(* IEC 61131-3 sources: daoli-st-library/DL_Device (part 10) *)

(* ---- FC_DL_RefSatPressToTemp.st ---- *)
(*
  ============================================================
  组件名 : FC_DL_RefSatPressToTemp
  分类   : DL_Device
  功能   : 制冷剂饱和压力转饱和温度，内置 R134a 与 R410A 分段线性表并做区间插值
  开源溯源 : internal-design（本轮无外部代码逐行引用）
             参考语义 : 无外部参考
  复杂度 : C2
  版本   : 1.0.0
  ============================================================
  表口径 : 压力为绝对压力 [bar abs]，温度为 [摄氏度]，两行表按 R134a 与 R410A 顺序平铺，
           行内压力严格升序；压力越出表范围时取端点温度并置 bValid 为假。
*)

FUNCTION FC_DL_RefSatPressToTemp : REAL
VAR_INPUT
    rPressBarA    : REAL; // 饱和绝对压力 [bar abs] saturation absolute pressure [bar abs]
    nRefrigerant  : INT; // 制冷剂 1=R134a 2=R410A [代号] refrigerant 1 for R134a and 2 for R410A [code]
END_VAR
VAR_OUTPUT
    rTempC : REAL; // 饱和温度 [摄氏度] saturation temperature [degree celsius]
    bValid : BOOL; // 结果有效标志 result validity flag
END_VAR
VAR CONSTANT
    afPress : ARRAY[0..1, 0..7] OF REAL := [1.0, 2.0, 4.0, 6.0, 8.0, 10.0, 14.0, 18.0, 1.0, 2.0, 4.0, 6.0, 8.0, 10.0, 14.0, 18.0]; // 饱和压力表 [bar abs] saturation pressure table [bar abs]
    afTemp  : ARRAY[0..1, 0..7] OF REAL := [-26.1, -10.1, 8.9, 21.6, 31.3, 39.4, 52.4, 62.5, -51.4, -34.1, -14.1, 0.4, 11.4, 20.5, 34.4, 45.0]; // 饱和温度表 [摄氏度] saturation temperature table [degree celsius]
    DL_IDX_LAST : INT := 7; // 表末下标 last table index
    DL_EPS_R    : REAL := 1.0E-6; // 实数零判定阈值 real zero threshold
END_VAR
VAR
    nRow  : INT := 0; // 表行号 0=R134a 1=R410A [行] table row number [row]
    nSeg  : INT := -1; // 命中区间下标，负为未命中 [段] hit segment index, negative when missing [segment]
    i     : INT := 0; // 区间游标 [段] segment cursor [segment]
    _rSpan: REAL := 0.0; // 区间压力跨度 [bar] segment pressure span [bar]
    _rFrac: REAL := 0.0; // 区间插值比例 [无量纲] interpolation fraction [dimensionless]
    _rT   : REAL := 0.0; // 温度中间量 [摄氏度] intermediate temperature [degree celsius]
END_VAR

// 段 1｜出口预置 preset the exit
FC_DL_RefSatPressToTemp := 0.0; // 缺省返回零 default zero return
rTempC := 0.0; // 温度预置零 temperature preset to zero
bValid := FALSE; // 计算完成前不认结果 unusable before the calculation
// 段 2｜非有限闸与制冷剂代号闸 finiteness gate and refrigerant code gate
IF (rPressBarA <> rPressBarA) OR (nRefrigerant < 1) OR (nRefrigerant > 2) THEN
    RETURN; // 非有限或代号非法即无效 non finite or an illegal code is void
END_IF
nRow := nRefrigerant - 1; // 行号由代号减一得出 the row index is the code minus one
// 段 3｜区间搜索 segment search over the ascending pressure table
FOR i := 0 TO (DL_IDX_LAST - 1) DO
    IF (rPressBarA >= afPress[nRow, i]) AND (rPressBarA <= afPress[nRow, i + 1]) THEN
        nSeg := i; // 命中升序区间 a segment is hit
    END_IF
END_FOR
// 段 4｜越界端点处理 endpoint handling for the out of table pressures
IF nSeg < 0 THEN
    IF rPressBarA < afPress[nRow, 0] THEN
        rTempC := afTemp[nRow, 0]; // 低于表底取表首温度 a pressure below the table takes the first temperature
    ELSE
        rTempC := afTemp[nRow, DL_IDX_LAST]; // 高于表顶取表末温度 a pressure above the table takes the last temperature
    END_IF
    RETURN; // 越界置无效并输出端点值 the out of table case is void with the endpoint emitted
END_IF
// 段 5｜线性插值 linear interpolation inside the hit segment
_rSpan := afPress[nRow, nSeg + 1] - afPress[nRow, nSeg]; // 区间压力跨度 segment pressure span
IF ABS(_rSpan) < DL_EPS_R THEN
    RETURN; // 跨度近零无法插值 a near zero span cannot interpolate
END_IF
_rFrac := (rPressBarA - afPress[nRow, nSeg]) / _rSpan; // 区间内插值比例 the fraction inside the segment
_rT := afTemp[nRow, nSeg] + _rFrac * (afTemp[nRow, nSeg + 1] - afTemp[nRow, nSeg]); // 端点温度线性插值 linear blend of the two temperatures
rTempC := _rT; // 温度落定 land the temperature
bValid := TRUE; // 结果可用 result usable
FC_DL_RefSatPressToTemp := _rT; // 函数返回饱和温度 return the saturation temperature
END_FUNCTION

(* ---- FC_DL_RefSatTempToPress.st ---- *)
(*
  ============================================================
  组件名 : FC_DL_RefSatTempToPress
  分类   : DL_Device
  功能   : 制冷剂饱和温度转饱和压力，内置 R134a 与 R410A 分段线性表并做区间插值
  开源溯源 : internal-design（本轮无外部代码逐行引用）
             参考语义 : 无外部参考
  复杂度 : C2
  版本   : 1.0.0
  ============================================================
  表口径 : 与压力查温度件同源的两张表，按温度升序重排后以温度为自变量插值压力；
           温度为绝对压力 [bar abs] 输出，温度越出表范围时取端点压力并置 bValid 为假。
*)

FUNCTION FC_DL_RefSatTempToPress : REAL
VAR_INPUT
    rTempC       : REAL; // 饱和温度 [摄氏度] saturation temperature [degree celsius]
    nRefrigerant : INT; // 制冷剂 1=R134a 2=R410A [代号] refrigerant 1 for R134a and 2 for R410A [code]
END_VAR
VAR_OUTPUT
    rPressBarA : REAL; // 饱和绝对压力 [bar abs] saturation absolute pressure [bar abs]
    bValid     : BOOL; // 结果有效标志 result validity flag
END_VAR
VAR CONSTANT
    afTemp  : ARRAY[0..1, 0..7] OF REAL := [-26.1, -10.1, 8.9, 21.6, 31.3, 39.4, 52.4, 62.5, -51.4, -34.1, -14.1, 0.4, 11.4, 20.5, 34.4, 45.0]; // 饱和温度表，行内升序 [摄氏度] saturation temperature table ascending inside each row [degree celsius]
    afPress : ARRAY[0..1, 0..7] OF REAL := [1.0, 2.0, 4.0, 6.0, 8.0, 10.0, 14.0, 18.0, 1.0, 2.0, 4.0, 6.0, 8.0, 10.0, 14.0, 18.0]; // 饱和压力表 [bar abs] saturation pressure table [bar abs]
    DL_IDX_LAST : INT := 7; // 表末下标 last table index
    DL_EPS_R    : REAL := 1.0E-6; // 实数零判定阈值 real zero threshold
END_VAR
VAR
    nRow  : INT := 0; // 表行号 0=R134a 1=R410A [行] table row number [row]
    nSeg  : INT := -1; // 命中区间下标，负为未命中 [段] hit segment index, negative when missing [segment]
    i     : INT := 0; // 区间游标 [段] segment cursor [segment]
    _rSpan: REAL := 0.0; // 区间温度跨度 [K] segment temperature span [kelvin]
    _rFrac: REAL := 0.0; // 区间插值比例 [无量纲] interpolation fraction [dimensionless]
    _rP   : REAL := 0.0; // 压力中间量 [bar abs] intermediate pressure [bar abs]
END_VAR

// 段 1｜出口预置 preset the exit
FC_DL_RefSatTempToPress := 0.0; // 缺省返回零 default zero return
rPressBarA := 0.0; // 压力预置零 pressure preset to zero
bValid := FALSE; // 计算完成前不认结果 unusable before the calculation
// 段 2｜非有限闸与制冷剂代号闸 finiteness gate and refrigerant code gate
IF (rTempC <> rTempC) OR (nRefrigerant < 1) OR (nRefrigerant > 2) THEN
    RETURN; // 非有限或代号非法即无效 non finite or an illegal code is void
END_IF
nRow := nRefrigerant - 1; // 行号由代号减一得出 the row index is the code minus one
// 段 3｜区间搜索 segment search over the ascending temperature table
FOR i := 0 TO (DL_IDX_LAST - 1) DO
    IF (rTempC >= afTemp[nRow, i]) AND (rTempC <= afTemp[nRow, i + 1]) THEN
        nSeg := i; // 命中升序区间 a segment is hit
    END_IF
END_FOR
// 段 4｜越界端点处理 endpoint handling for the out of table temperatures
IF nSeg < 0 THEN
    IF rTempC < afTemp[nRow, 0] THEN
        rPressBarA := afPress[nRow, 0]; // 低于表底取表首压力 a temperature below the table takes the first pressure
    ELSE
        rPressBarA := afPress[nRow, DL_IDX_LAST]; // 高于表顶取表末压力 a temperature above the table takes the last pressure
    END_IF
    RETURN; // 越界置无效并输出端点值 the out of table case is void with the endpoint emitted
END_IF
// 段 5｜线性插值 linear interpolation inside the hit segment
_rSpan := afTemp[nRow, nSeg + 1] - afTemp[nRow, nSeg]; // 区间温度跨度 segment temperature span
IF ABS(_rSpan) < DL_EPS_R THEN
    RETURN; // 跨度近零无法插值 a near zero span cannot interpolate
END_IF
_rFrac := (rTempC - afTemp[nRow, nSeg]) / _rSpan; // 区间内插值比例 the fraction inside the segment
_rP := afPress[nRow, nSeg] + _rFrac * (afPress[nRow, nSeg + 1] - afPress[nRow, nSeg]); // 端点压力线性插值 linear blend of the two pressures
rPressBarA := _rP; // 压力落定 land the pressure
bValid := TRUE; // 结果可用 result usable
FC_DL_RefSatTempToPress := _rP; // 函数返回饱和压力 return the saturation pressure
END_FUNCTION

(* ---- FC_DL_RefSubcoolCalc.st ---- *)
(*
  ============================================================
  组件名 : FC_DL_RefSubcoolCalc
  分类   : DL_Device
  功能   : 液管过冷度计算，由冷凝饱和温度与液管温度求过冷度并分档判定
  开源溯源 : internal-design（本轮无外部代码逐行引用）
             参考语义 : 无外部参考
  复杂度 : C1
  版本   : 1.0.0
  ============================================================
*)

FUNCTION FC_DL_RefSubcoolCalc : REAL
VAR_INPUT
    rLiquidTempC    : REAL; // 液管实测温度 [摄氏度] measured liquid line temperature [degree celsius]
    rSatLiquidTempC : REAL; // 液管饱和温度 [摄氏度] saturation temperature at the liquid pressure [degree celsius]
    rScLow          : REAL; // 过冷度下限 [K] lower subcooling bound [kelvin]
    rScHigh         : REAL; // 过冷度上限 [K] upper subcooling bound [kelvin]
END_VAR
VAR_OUTPUT
    rSubcoolK : REAL; // 液管过冷度 [K] liquid subcooling [kelvin]
    nStatus   : INT; // 分档 0正常 1偏低 2偏高 [档] status 0 normal, 1 low, 2 high [band]
    bValid    : BOOL; // 结果有效标志 result validity flag
END_VAR
VAR
    _bFin  : BOOL := FALSE; // 四输入有限性判定 finiteness verdict of the four inputs
    _rSc   : REAL := 0.0; // 过冷度中间量 [K] intermediate subcooling [kelvin]
    _rLo   : REAL := 0.0; // 钳位后的下限 [K] clamped lower bound [kelvin]
    _rHi   : REAL := 0.0; // 钳位后的上限 [K] clamped upper bound [kelvin]
END_VAR

// 段 1｜出口预置 preset the exit
FC_DL_RefSubcoolCalc := 0.0; // 缺省返回零 default zero return
rSubcoolK := 0.0; // 过冷度预置零 subcooling preset to zero
nStatus := 0; // 分档预置正常 status preset normal
bValid := FALSE; // 计算完成前不认结果 unusable before the calculation
// 段 2｜非有限闸 finiteness gate
_bFin := (rLiquidTempC = rLiquidTempC) AND (rSatLiquidTempC = rSatLiquidTempC) AND (rScLow = rScLow) AND (rScHigh = rScHigh); // 四输入自反判定 self comparison of the four inputs
IF NOT _bFin THEN
    RETURN; // 非有限即无效 non finite means invalid
END_IF
// 段 3｜主体过冷度 main subcooling，口径为饱和温度减液管温度 saturation minus the liquid temperature
_rSc := rSatLiquidTempC - rLiquidTempC; // 饱和温度减液管温度 saturation minus the liquid temperature
rSubcoolK := _rSc; // 过冷度落定 land the subcooling
// 段 4｜上下限整形 bound reshape
_rLo := rScLow; // 取下限 take the lower bound
_rHi := rScHigh; // 取上限 take the upper bound
IF _rLo > _rHi THEN
    _rLo := rScHigh; // 上下限倒置时下限取原上限 an inverted pair swaps the lower bound
    _rHi := rScLow; // 上下限倒置时上限取原下限 an inverted pair swaps the upper bound
END_IF
// 段 5｜双向分档判定 directional status verdict
IF _rSc < _rLo THEN
    nStatus := 1; // 过冷度偏低 subcooling too low
ELSIF _rSc > _rHi THEN
    nStatus := 2; // 过冷度偏高 subcooling too high
ELSE
    nStatus := 0; // 区间内正常 inside the normal band
END_IF
bValid := TRUE; // 结果可用 result usable
FC_DL_RefSubcoolCalc := _rSc; // 函数返回过冷度 return the subcooling
END_FUNCTION

(* ---- FC_DL_RefSuperheatCalc.st ---- *)
(*
  ============================================================
  组件名 : FC_DL_RefSuperheatCalc
  分类   : DL_Device
  功能   : 吸气过热度计算，由吸气温度与对应饱和温度求过热度并分档判定
  开源溯源 : internal-design（本轮无外部代码逐行引用）
             参考语义 : 无外部参考
  复杂度 : C1
  版本   : 1.0.0
  ============================================================
*)

FUNCTION FC_DL_RefSuperheatCalc : REAL
VAR_INPUT
    rSuctionTempC    : REAL; // 吸气实测温度 [摄氏度] measured suction temperature [degree celsius]
    rSatSuctionTempC : REAL; // 吸气饱和温度 [摄氏度] saturation temperature at the suction pressure [degree celsius]
    rShLow           : REAL; // 过热度下限 [K] lower superheat bound [kelvin]
    rShHigh          : REAL; // 过热度上限 [K] upper superheat bound [kelvin]
END_VAR
VAR_OUTPUT
    rSuperheatK : REAL; // 吸气过热度 [K] suction superheat [kelvin]
    nStatus     : INT; // 分档 0正常 1偏低 2偏高 [档] status 0 normal, 1 low, 2 high [band]
    bValid      : BOOL; // 结果有效标志 result validity flag
END_VAR
VAR
    _bFin  : BOOL := FALSE; // 四输入有限性判定 finiteness verdict of the four inputs
    _rSh   : REAL := 0.0; // 过热度中间量 [K] intermediate superheat [kelvin]
    _rLo   : REAL := 0.0; // 钳位后的下限 [K] clamped lower bound [kelvin]
    _rHi   : REAL := 0.0; // 钳位后的上限 [K] clamped upper bound [kelvin]
END_VAR

// 段 1｜出口预置 preset the exit
FC_DL_RefSuperheatCalc := 0.0; // 缺省返回零 default zero return
rSuperheatK := 0.0; // 过热度预置零 superheat preset to zero
nStatus := 0; // 分档预置正常 status preset normal
bValid := FALSE; // 计算完成前不认结果 unusable before the calculation
// 段 2｜非有限闸 finiteness gate
_bFin := (rSuctionTempC = rSuctionTempC) AND (rSatSuctionTempC = rSatSuctionTempC) AND (rShLow = rShLow) AND (rShHigh = rShHigh); // 四输入自反判定 self comparison of the four inputs
IF NOT _bFin THEN
    RETURN; // 非有限即无效 non finite means invalid
END_IF
// 段 3｜主体过热度 main superheat
_rSh := rSuctionTempC - rSatSuctionTempC; // 吸气温度减饱和温度 suction minus saturation
rSuperheatK := _rSh; // 过热度落定 land the superheat
// 段 4｜上下限整形 bound reshape
_rLo := rShLow; // 取下限 take the lower bound
_rHi := rShHigh; // 取上限 take the upper bound
IF _rLo > _rHi THEN
    _rLo := rShHigh; // 上下限倒置时下限取原上限 an inverted pair swaps the lower bound
    _rHi := rShLow; // 上下限倒置时上限取原下限 an inverted pair swaps the upper bound
END_IF
// 段 5｜双向分档判定 directional status verdict
IF _rSh < _rLo THEN
    nStatus := 1; // 过热度偏低 superheat too low
ELSIF _rSh > _rHi THEN
    nStatus := 2; // 过热度偏高 superheat too high
ELSE
    nStatus := 0; // 区间内正常 inside the normal band
END_IF
bValid := TRUE; // 结果可用 result usable
FC_DL_RefSuperheatCalc := _rSh; // 函数返回过热度 return the superheat
END_FUNCTION

(* ---- FC_DL_SheetPeelForceCalc.st ---- *)
(*
  ============================================================
  组件名 : FC_DL_SheetPeelForceCalc
  分类   : DL_Device
  功能   : 片材剥离力计算，由接触面积粘附强度与静电电压求剥离力并按剥离角折减
  复杂度 : C2
  版本   : 1.0.0
  作者   : 道莅工业代码库工厂 / R81
  日期   : 2026-11-24
  开源溯源 : clean-room（no upstream）—— 依据公开工程公式自研，未复制任何上游实现
  红线自检 : R1 无GVL/R2 无物理地址/R3 纯IEC/R4 防除零/R5 双语注释
  接口说明 :
      粘附分量 = 接触面积(m2) * 粘附强度(Pa)，面积由 mm2 乘 1e-6，强度由 kPa 乘 1000。
      静电分量 = 静电电压(kV) * 0.05，系数为工程经验折算，单位 N/kV。
      剥离角修正系数 = (1 + COS(角度)) / 2，归一到 0 度时为 1、90 度为 0.5、180 度为 0，便于跨机型比较。
      剥离力超过 50 N 判需要外部辅助剥离。
  ============================================================
*)
FUNCTION FC_DL_SheetPeelForceCalc : BOOL
VAR_INPUT
    bEnable       : BOOL; // 使能：TRUE 时计算 / Enable: TRUE to compute
    bErr          : BOOL; // 外部故障：TRUE 时立即退出并置结果无效 / External fault: TRUE aborts with invalid result
    rArea_mm2     : REAL; // 片材与承载面接触面积 [mm2] / contact area between sheet and support [square millimetre]
    rAdhesion_kpa : REAL; // 单位面积粘附强度 [kPa] / adhesion strength per unit area [kilopascal]
    rStaticKv     : REAL; // 片材静电电位 [kV] / electrostatic potential of the sheet [kilovolt]
    rPeelAngleDeg : REAL; // 剥离角度，0 度表示垂直拉起 [度] / peel angle, zero means lifting perpendicular [degree]
END_VAR
VAR_OUTPUT
    rAdhesionN : REAL; // 粘附力分量 [N] / adhesion force component [newton]
    rStaticN   : REAL; // 静电力分量 [N] / electrostatic force component [newton]
    rAngleFactor : REAL; // 剥离角折减系数，0~1 [无量纲] / peel angle reduction factor from 0 to 1 [dimensionless]
    rPeelN     : REAL; // 综合剥离力 [N] / resultant peel force [newton]
    bNeedAssist : BOOL; // 需要辅助：TRUE 表示剥离力超过 50 N / assistance required, TRUE when the peel force exceeds 50 newton
    bValid     : BOOL; // 输出有效：TRUE 表示结果可用 / Output valid
END_VAR
VAR CONSTANT
    DL_R_MAX     : REAL := 3.0E38;     // 实数上界，用于拦截 Inf [无量纲] / real upper bound used to reject infinity [dimensionless]
    DL_EPS       : REAL := 1.0E-12;    // 除零判定阈值 [无量纲] / division guard threshold [dimensionless]
    DL_MM2_TO_M2 : REAL := 1.0E-6;     // 平方毫米折平方米系数 [m2/mm2] / square millimetre to square metre factor [square metre per square millimetre]
    DL_KPA_TO_PA : REAL := 1000.0;     // 千帕折帕系数 [Pa/kPa] / kilopascal to pascal factor [pascal per kilopascal]
    DL_KV_TO_N   : REAL := 0.05;       // 每千伏静电折算力 [N/kV] / electrostatic force per kilovolt [newton per kilovolt]
    DL_DEG_TO_RAD : REAL := 0.0174533; // 度转弧度系数 [rad/度] / degree to radian factor [radian per degree]
    DL_HALF      : REAL := 0.5;        // 二分之一，用于角度系数归一 [无量纲] / one half used to normalise the angle factor [dimensionless]
    DL_ONE       : REAL := 1.0;        // 单位常量 [无量纲] / unity constant [dimensionless]
    DL_ASSIST_N  : REAL := 50.0;       // 辅助剥离门限 [N] / assistance threshold [newton]
    DL_ANGLE_MAX : REAL := 180.0;      // 剥离角允许上限 [度] / permitted upper bound of the peel angle [degree]
    DL_STAT_MAX  : REAL := 1000.0;     // 静电电位合理上限 [kV] / sanity upper bound of the electrostatic potential [kilovolt]
END_VAR
VAR
    _bFin  : BOOL := FALSE; // 输入有限性判定结果 / input finiteness verdict
    _rRad  : REAL := 0.0;   // 剥离角折算弧度 [rad] / peel angle in radian [radian]
END_VAR

    // 段 1｜出口预置
    rAdhesionN := 0.0;
    rStaticN := 0.0;
    rAngleFactor := 0.0;
    rPeelN := 0.0;
    bNeedAssist := FALSE;
    bValid := FALSE;
    // 段 2｜使能闸与外部故障闸
    IF NOT bEnable THEN
        RETURN;
    END_IF;
    IF bErr THEN
        RETURN;
    END_IF;
    // 段 3｜非有限闸
    _bFin := (rArea_mm2 = rArea_mm2) AND (ABS(rArea_mm2) <= DL_R_MAX) AND (rAdhesion_kpa = rAdhesion_kpa) AND (ABS(rAdhesion_kpa) <= DL_R_MAX) AND (rStaticKv = rStaticKv) AND (ABS(rStaticKv) <= DL_R_MAX) AND (rPeelAngleDeg = rPeelAngleDeg) AND (ABS(rPeelAngleDeg) <= DL_R_MAX);
    IF NOT _bFin THEN
        RETURN;
    END_IF;
    // 段 4｜域闸：面积非负、粘附强度非负、静电位非负且合理、角度 0~180
    IF (rArea_mm2 < 0.0) OR (rAdhesion_kpa < 0.0) OR (rStaticKv < 0.0) OR (rStaticKv > DL_STAT_MAX) THEN
        RETURN;
    END_IF;
    IF (rPeelAngleDeg < 0.0) OR (rPeelAngleDeg > DL_ANGLE_MAX) THEN
        RETURN;
    END_IF;
    // 段 5｜两个力分量
    rAdhesionN := rArea_mm2 * DL_MM2_TO_M2 * rAdhesion_kpa * DL_KPA_TO_PA;
    rStaticN := rStaticKv * DL_KV_TO_N;
    // 段 6｜角度折减系数
    _rRad := rPeelAngleDeg * DL_DEG_TO_RAD;
    rAngleFactor := (DL_ONE + COS(_rRad)) * DL_HALF;
    IF rAngleFactor < 0.0 THEN
        rAngleFactor := 0.0;
    END_IF;
    IF rAngleFactor > DL_ONE THEN
        rAngleFactor := DL_ONE;
    END_IF;
    // 段 7｜综合剥离力
    rPeelN := (rAdhesionN + rStaticN) * rAngleFactor;
    // 段 8｜辅助判定
    IF rPeelN > DL_ASSIST_N THEN
        bNeedAssist := TRUE;
    ELSE
        bNeedAssist := FALSE;
    END_IF;
    bValid := TRUE;
    FC_DL_SheetPeelForceCalc := bValid;
END_FUNCTION

(* ---- FC_DL_SizeApplicatorPickupCalc.st ---- *)
// FC_DL_SizeApplicatorPickupCalc v1.0.0
// 开源溯源：clean-room 自研（族 DL_Device，ST 生态实测 0 命中，无外部代码引入）
(*
  功能: 上胶率：干基量 = 浸润剂流量·固含量/100 [kg/h]（乳液密度按 1.0 kg/L，L/h 数值等同 kg/h），
        上胶率 = 100·干基量/丝束产出 [%]。
  邻件/码位: 与 FC_DL_StrandTensionAtWinderCalc 同属拉丝后端条件件（化学上胶 vs 力学张力）；
             16#0002_9225 = 非有限、产出非正、流量为负、固含量越界或上胶率出 0.1~3.0%。
*)
FUNCTION FC_DL_SizeApplicatorPickupCalc : REAL
VAR_INPUT
    fSizeFlow   : REAL := 40.0;     // 浸润剂流量 [L/h]，域 >= 0 / Size flow [L/h]
    fSizeSolids : REAL := 6.0;      // 固含量 [%]，域 (0, 100] / Solids content [%]
    fStrandRate : REAL := 120.0;    // 丝束产出 [kg/h]，域 > 0 / Strand output [kg/h]
END_VAR
VAR_OUTPUT
    fPickup  : REAL;                // 上胶率 [%]，工艺窗 0.1~3.0 / Size pickup [%]
    bValid   : BOOL;                // 结果有效回执 [-] / Result validity receipt
    uErrorId : UDINT;               // 事件码，0 = 无事件 / Event code
END_VAR
VAR
    fDryBasis : REAL := 0.0;        // 干基上胶量 [kg/h] / Dry size basis [kg/h]
END_VAR
// 段 0：全路径出口安全缺省 / Safe defaults on all outlets
fPickup := 0.0;                 // 上胶率缺省零 / Pickup default zero
bValid := FALSE;                // 有效回执预清 / Validity preset clear
uErrorId := 16#0000;            // 事件码预清 / Event code preset clear
FC_DL_SizeApplicatorPickupCalc := 0.0;  // 返回值缺省零（镜像上胶率）/ Return default zero
// 段 1：非有限闸（三入参全枚举）/ Non-finite gate over all inputs
IF (fSizeFlow <> fSizeFlow) OR (fSizeSolids <> fSizeSolids) OR (fStrandRate <> fStrandRate)
   OR (ABS(fSizeFlow) >= 3.0E38) OR (ABS(fSizeSolids) >= 3.0E38) OR (ABS(fStrandRate) >= 3.0E38) THEN
    uErrorId := 16#0002_9225;   // 入参非有限拒收 / Non-finite input reject
    RETURN;
END_IF
// 段 2：域闸（产出为正防除零 + 流量非负 + 固含量区间，R4）/ Domain gate
IF fStrandRate <= 1.0E-6 THEN
    uErrorId := 16#0002_9225;   // 丝束产出非正，上胶率不可解 / Non-positive strand rate
    RETURN;
END_IF
IF fSizeFlow < 0.0 THEN
    uErrorId := 16#0002_9225;   // 流量为负 / Negative flow
    RETURN;
END_IF
IF (fSizeSolids <= 0.0) OR (fSizeSolids > 100.0) THEN
    uErrorId := 16#0002_9225;   // 固含量越界 / Solids content out of range
    RETURN;
END_IF
// 段 3：主计算（干基量 → 上胶率）/ Main computation
fDryBasis := fSizeFlow * fSizeSolids / 100.0;                   // 干基量 [kg/h] / Dry basis
fPickup := 100.0 * fDryBasis / fStrandRate;                     // 上胶率 [%] / Size pickup
// 段 4：出口闸（非有限复核 + 0.1~3.0% 工艺窗判定）/ Outlet gate
IF (fPickup <> fPickup) OR (ABS(fPickup) >= 3.0E38) OR (fPickup < 0.0) THEN
    fPickup := 0.0;             // 复核失败回缺省 / Fallback on recheck failure
    uErrorId := 16#0002_9225;   // 出口复核拒收 / Output recheck reject
    RETURN;
END_IF
IF (fPickup < 0.1) OR (fPickup > 3.0) THEN
    uErrorId := 16#0002_9225;   // 信息级：上胶率出工艺窗 / Info: pickup out of window
    RETURN;                     // bValid 保持 FALSE / Validity stays false
END_IF
bValid := TRUE;                 // 有效回执 / Validity receipt
FC_DL_SizeApplicatorPickupCalc := fPickup;      // 返回值镜像上胶率 / Return mirrors pickup
END_FUNCTION

(* ---- FC_DL_SlitterKnifeClearanceCalc.st ---- *)
(*
  Name: FC_DL_SlitterKnifeClearanceCalc
  Category: DL_Device
  Version: 1.0.0
  Round: R89 / 2026-11-25
  开源溯源：clean-room 自研（族 板带剪切分条卷取，ST 开源生态实测 0 命中，无外部代码引入）
  功能：分条圆盘刀侧间隙与刀盘重叠量：基准间隙率随抗拉强度线性修正后乘厚度。
  边界条件：① 三入参全部过非有限闸，任一非有限返回哨兵 -1；
            ② 间隙率修正以 400 MPa 为基准点、每 100 MPa 增减 0.5 个百分点，修正后钳位 2~14 %；
            ③ 重叠量取侧间隙的 15 %（薄料防刀口顶死经验值），随间隙同比缩放，无量纲系数见常量；
            ④ 钳位属量值饱和，置 xValid 保持 TRUE（厚度与强度均已合法）。
  量纲自证：pct[%]/100 无量纲；thk[mm] × 无量纲 = mm。
*)
FUNCTION FC_DL_SlitterKnifeClearanceCalc : REAL
VAR_INPUT
    fThkMm : REAL;          (* 带钢厚度 [mm] Strip thickness [mm] *)
    fTensileMpa : REAL;     (* 抗拉强度 [MPa] Tensile strength [MPa] *)
    fClearPctBase : REAL;   (* 基准间隙率（400 MPa 基准点） [%] Base clearance ratio at 400 MPa [%] *)
END_VAR
VAR_OUTPUT
    fClearanceMm : REAL;    (* 侧间隙 [mm] Side clearance [mm] *)
    fOverlapMm : REAL;      (* 刀盘重叠量 [mm] Knife overlap [mm] *)
    xValid : BOOL;          (* 计算有效性标志 [-] Calculation valid flag *)
END_VAR
VAR CONSTANT
    DL_KNIFE_TSREF : REAL := 400.0;     (* 间隙率基准强度 [MPa] Reference tensile strength [MPa] *)
    DL_KNIFE_SLOPE : REAL := 0.5;       (* 每 100 MPa 间隙率增量 [%/100MPa] Ratio increment per 100 MPa *)
    DL_KNIFE_OVL : REAL := 0.15;        (* 重叠量/侧间隙比 [-] Overlap to clearance ratio *)
    DL_KNIFE_PCT_LO : REAL := 2.0;      (* 间隙率下限 [%] Clearance ratio floor [%] *)
    DL_KNIFE_PCT_HI : REAL := 14.0;     (* 间隙率上限 [%] Clearance ratio ceiling [%] *)
    DL_PCT : REAL := 100.0;             (* 百分数基准 [%] Percent base *)
    DL_T_MIN : REAL := 0.1;             (* 带厚下限 [mm] Thickness floor [mm] *)
    DL_T_MAX : REAL := 6.0;             (* 带厚上限 [mm] Thickness ceiling [mm] *)
    DL_TS_MIN : REAL := 200.0;          (* 强度下限 [MPa] Tensile floor [MPa] *)
    DL_TS_MAX : REAL := 1500.0;         (* 强度上限 [MPa] Tensile ceiling [MPa] *)
    DL_B_MIN : REAL := 1.0;             (* 基准间隙率下限 [%] Base ratio floor [%] *)
    DL_B_MAX : REAL := 15.0;            (* 基准间隙率上限 [%] Base ratio ceiling [%] *)
END_VAR
VAR
    fPct : REAL;    (* 修正后间隙率 [%] Corrected clearance ratio [%] *)
END_VAR
(* 出口预置：三出口统一预置（R256） *)
fClearanceMm := 0.0; fOverlapMm := 0.0; xValid := FALSE;
(* 非有限闸：NaN 自反判 + Inf 差值自减判，三入参全枚举 *)
IF (fThkMm <> fThkMm) OR ((fThkMm - fThkMm) <> 0.0)
   OR (fTensileMpa <> fTensileMpa) OR ((fTensileMpa - fTensileMpa) <> 0.0)
   OR (fClearPctBase <> fClearPctBase) OR ((fClearPctBase - fClearPctBase) <> 0.0) THEN
    FC_DL_SlitterKnifeClearanceCalc := -1.0;    (* 哨兵 -1：入参非有限 / Sentinel -1, non-finite input *)
    RETURN;
END_IF
(* 组态域闸：厚度、强度、基准间隙率逐项定域 *)
IF (fThkMm < DL_T_MIN) OR (fThkMm > DL_T_MAX)
   OR (fTensileMpa < DL_TS_MIN) OR (fTensileMpa > DL_TS_MAX)
   OR (fClearPctBase < DL_B_MIN) OR (fClearPctBase > DL_B_MAX) THEN
    FC_DL_SlitterKnifeClearanceCalc := -1.0;    (* 哨兵 -1：组态非法 / Sentinel -1, bad configuration *)
    RETURN;
END_IF
(* 强度线性修正：pct = base + slope·(σ − σref)/100，斜率单位 %/100MPa *)
fPct := fClearPctBase + DL_KNIFE_SLOPE * ((fTensileMpa - DL_KNIFE_TSREF) / DL_PCT);
(* 修正后钳位：低于下限刀口挤压、高于上限毛刺超差 *)
IF fPct < DL_KNIFE_PCT_LO THEN
    fPct := DL_KNIFE_PCT_LO;
ELSIF fPct > DL_KNIFE_PCT_HI THEN
    fPct := DL_KNIFE_PCT_HI;
END_IF
(* 侧间隙：thk[mm] × pct[%]/100 = mm *)
fClearanceMm := fThkMm * (fPct / DL_PCT);
(* 重叠量：侧间隙 × 经验比，无量纲系数，量纲保持 mm *)
fOverlapMm := fClearanceMm * DL_KNIFE_OVL;
xValid := TRUE;                                 (* 链路有效 / Chain valid *)
FC_DL_SlitterKnifeClearanceCalc := fClearanceMm;
END_FUNCTION

(* ---- FC_DL_SlotHeightFitCalc.st ---- *)
(*
  DL Factory R83 | FC_DL_SlotHeightFitCalc
  功能：校验货位净高对托盘货高的容纳能力，给出净余量与高度利用率。
  开源溯源：无（clean-room 自研，依据公开工艺公式，来源=行业通用公式，许可证=MIT，借鉴点=公式结构）
  规则：R1-R21 全遵守
*)
FUNCTION FC_DL_SlotHeightFitCalc : REAL
VAR_INPUT
    fSlotClearHmm  : REAL; // 货位净高（横梁下沿到地面）[mm] / Slot clear height [mm]
    fPalletHmm     : REAL; // 托盘货高（含托盘本体）[mm] / Pallet load height incl. pallet [mm]
    fLiftClearMm   : REAL; // 存取所需起升余量 [mm] / Required lift clearance [mm]
    fTolMm         : REAL; // 允许最小安全余量 [mm] / Required minimum safety margin [mm]
END_VAR
VAR_OUTPUT
    fMarginMm : REAL; // 净余量（净高-货高-起升余量）[mm] / Net margin [mm]
    fUtilPct  : REAL; // 高度利用率（货高÷净高）[%] / Height utilisation [%]
    xFit      : BOOL; // 匹配判定（余量不低于安全余量）/ Fit decision
    xValid    : BOOL; // 计算有效性标志 / Calculation validity flag
END_VAR

// ---------- 输出预置 ----------
fMarginMm := 0.0;                   // 余量清零 [mm] / Margin zeroed
fUtilPct  := 0.0;                   // 利用率清零 [%] / Utilisation zeroed
xFit      := FALSE;                 // 预置不匹配（安全侧）/ Preset no-fit (safe side)
xValid    := FALSE;                 // 有效性预置 FALSE / Validity preset FALSE

// ---------- 非有限拦截 + 量纲自检（R20/R21） ----------
IF NOT (fSlotClearHmm > -1.0E30 AND fSlotClearHmm < 1.0E30) OR NOT (fPalletHmm > -1.0E30 AND fPalletHmm < 1.0E30) OR NOT (fLiftClearMm > -1.0E30 AND fLiftClearMm < 1.0E30) OR NOT (fTolMm > -1.0E30 AND fTolMm < 1.0E30) OR fSlotClearHmm <= 0.0 OR fPalletHmm <= 0.0 OR fLiftClearMm < 0.0 OR fTolMm < 0.0 THEN
    FC_DL_SlotHeightFitCalc := -1.0; // 哨兵 -1：非有限或量纲越界 / Sentinel -1: non-finite or out of domain
    RETURN;
END_IF

// ---------- 净余量：同量纲相减（mm），三件均以 mm 输入故无需换算 ----------
fMarginMm := fSlotClearHmm - fPalletHmm - fLiftClearMm; // 净余量 [mm] / Net margin [mm]

// ---------- 高度利用率：货高 ÷ 净高 × 100，净高分母显式零闸（R4/R21） ----------
IF ABS(fSlotClearHmm) > 1.0E-9 THEN               // 净高分母显式零闸 / Explicit zero gate on clear height
    fUtilPct := (fPalletHmm / fSlotClearHmm) * 100.0; // 高度利用率 [%] / Height utilisation [%]
ELSE
    fUtilPct := 0.0;                // 除零防御缺省 [%] / Divide-by-zero default
END_IF

// ---------- 匹配判定：余量不低于安全余量（单一比较，禁浮点等号） ----------
xFit   := fMarginMm >= fTolMm;      // 匹配布尔 / Fit boolean
xValid := TRUE;                     // 链路有效 / Chain valid
FC_DL_SlotHeightFitCalc := fMarginMm; // 返回净余量 [mm] / Return net margin [mm]
END_FUNCTION

(* ---- FC_DL_SodiumPnaCalc.st ---- *)
(* ============================================================
   DL_Device / FC_DL_SodiumPnaCalc ｜ v1.0.0 ｜ 2026-11-25
   功能：钠离子 pNa 换算 pNa = (0 − E_mv) / S(T) [−]，S(T) = S25 · (273.15 + T) / 298.15
         [mV/decade]；内部按 [Na] = 23 g/mol 折算 µg/L = 23 · 10^(6 − pNa) 用于量程判据。
   边界：斜率 ≤ 0 或温度越出 [−5, 80]°C → 钳定后仍不可解：pNa 写 0、bOutOfRange=TRUE；
         任一入参非有限 → pNa 写 0、bOutOfRange=TRUE（N1 安全侧）；
         nSlopeSel：0=理论斜率 59.16，1=实测钠电极斜率 56.0，其余按理论斜率并
         判为量程外（档位非法）。签名只有一个 REAL 出口，故 pNa 为主出口，
         µg/L 仅在内部参与量程判据（本件相对规划的收窄点，不改签名）。
         量纲清单（N5）：1 mol/L NaCl = 23 g/L；1 mg/L = 1000 µg/L；
         量程 0.1 ~ 100000 µg/L ↔ pNa 8.36 ~ 2.36。
   依赖：仅 IEC 61131-3（EXPT / ABS） ｜ 溯源：DLF-D-WATERANA
   验收：mV=−325、T=25、档位 0 → S=59.16 → pNa≈5.494、未越限；
         档位 1 → S=56.0 → pNa≈5.804；斜率不可解 → pNa=0、越限。
   ============================================================ *)
FUNCTION FC_DL_SodiumPnaCalc : BOOL
VAR_INPUT
    fMvMeas   : REAL;  // 钠电极实测电位 [mV] / Measured sodium electrode potential
    fTempC    : REAL;  // 水样温度 [°C] / Sample temperature in Celsius degrees
    nSlopeSel : INT;   // 斜率档位 0=理论 1=实测钠电极 [-] / Slope selector
END_VAR
VAR_OUTPUT
    fPna        : REAL;  // 钠离子 pNa 值 [-] / Sodium pNa value
    bOutOfRange : BOOL;  // pNa 越出测量量程或输入非法 [-] / pNa outside the measurement range or illegal input
END_VAR
VAR
    _fT     : REAL;  // 钳定后温度 [°C] / Clamped temperature
    _fS25   : REAL;  // 25°C 下的斜率基值 [mV/decade] / Slope base at twenty five Celsius
    _fSlope : REAL;  // 温度修正后斜率 [mV/decade] / Temperature corrected slope
    _fPna   : REAL;  // pNa 中间值 [-] / Intermediate pNa value
    _fUgL   : REAL;  // 折算钠浓度 [µg/L] / Converted sodium concentration
    _bBad   : BOOL;  // 输入或档位非法标志 [-] / Illegal input or selector flag
END_VAR
VAR CONSTANT
    DL_SOD_S25  : REAL := 59.16;    // 25 摄氏度理论斜率 [mV/decade] / Theoretical slope at twenty five Celsius
    DL_SOD_S56  : REAL := 56.0;     // 实测钠电极斜率（25°C）[mV/decade] / Measured sodium electrode slope
    DL_SOD_TREF : REAL := 25.0;     // 参考温度 [°C] / Reference temperature
    DL_SOD_TK   : REAL := 273.15;   // 绝对零度偏移 [K] / Kelvin offset of the Celsius scale
    DL_SOD_TLO  : REAL := -5.0;     // 温度域下限 [°C] / Lower temperature bound
    DL_SOD_THI  : REAL := 80.0;     // 温度域上限 [°C] / Upper temperature bound
    DL_SOD_MOL  : REAL := 23.0;     // 钠摩尔质量 [g/mol] / Molar mass of sodium
    DL_SOD_UGLO : REAL := 0.1;      // 折算浓度下限 [µg/L] / Lower bound of the converted concentration
    DL_SOD_UGHI : REAL := 100000.0; // 折算浓度上限 [µg/L] / Upper bound of the converted concentration
    DL_SOD_DEC  : REAL := 6.0;      // pNa → µg/L 的十进制移位 [-] / Decade shift from pNa to micrograms per liter
END_VAR

(* 段 0：出口预置安全侧（pNa 0、越限置位，N1/N3） *)
FC_DL_SodiumPnaCalc := FALSE;
fPna := 0.0;  bOutOfRange := TRUE;
_bBad := FALSE;

(* 段 1：非有限闸（两个浮点入参） *)
IF (fMvMeas <> fMvMeas) OR (fTempC <> fTempC) THEN RETURN; END_IF

(* 段 2：温度域闸（越域钳定并判为越限，禁外推） *)
_fT := fTempC;
IF fTempC < DL_SOD_TLO THEN
    _fT := DL_SOD_TLO;  _bBad := TRUE;
ELSIF fTempC > DL_SOD_THI THEN
    _fT := DL_SOD_THI;  _bBad := TRUE;
END_IF

(* 段 3：斜率分派（非法档位按理论斜率并判越限） *)
CASE nSlopeSel OF
0:      _fS25 := DL_SOD_S25;
1:      _fS25 := DL_SOD_S56;
ELSE
    _fS25 := DL_SOD_S25;  _bBad := TRUE;
END_CASE
_fSlope := _fS25 * (_fT + DL_SOD_TK) / (DL_SOD_TREF + DL_SOD_TK);

(* 段 4：pNa 与折算浓度（除子已证 > 0，S25 恒为正） *)
IF _fSlope <= 0.0 THEN RETURN; END_IF
_fPna := (0.0 - fMvMeas) / _fSlope;
IF (_fPna <> _fPna) OR ((_fPna - _fPna) <> (_fPna - _fPna)) THEN RETURN; END_IF
_fUgL := DL_SOD_MOL * EXPT(10.0, DL_SOD_DEC - _fPna);

(* 段 5：单一出口裁决（判据与出口同源于 _fPna/_fUgL，N4/R23） *)
IF _bBad OR (_fUgL <> _fUgL) OR ((_fUgL - _fUgL) <> (_fUgL - _fUgL)) THEN
    fPna := 0.0;                        // 非有限或组态非法：落安全侧
    bOutOfRange := TRUE;
    RETURN;
END_IF
IF (_fUgL < DL_SOD_UGLO) OR (_fUgL > DL_SOD_UGHI) THEN
    fPna := _fPna;                      // 出量程：值照给供上层记录
    bOutOfRange := TRUE;
    RETURN;
END_IF
fPna := _fPna;
bOutOfRange := FALSE;
FC_DL_SodiumPnaCalc := TRUE;
END_FUNCTION

(* ---- FC_DL_SpareReorderPoint.st ---- *)
(*
  道莅工业代码库 / Daoli Industrial ST Library
  组件: FC_DL_SpareReorderPoint
  分类: DL_Device
  开源溯源: 无（clean-room 工程公式自研；参考公开工艺计算公式，未复制任何受版权保护代码）
  许可证: 本项目自有 (MIT)
  功能: 备件订货点与缺料量计算，触发补货判定
*)
FUNCTION FC_DL_SpareReorderPoint : BOOL
VAR_INPUT
    rDailyUse : REAL; // 日均消耗量 [件/d] / average daily consumption
    rLeadDays : REAL; // 采购提前期 [d] / procurement lead time in days
    rSafetyDays : REAL; // 安全库存天数 [d] / safety stock in days
    rOnHand : REAL; // 当前在手库存 [件] / stock on hand
END_VAR
VAR_OUTPUT
    rRop : REAL; // 订货点 [件] / reorder point
    rShortQty : REAL; // 相对订货点的缺口量 [件] / shortage against the reorder point
    bValid : BOOL; // 结果有效位 [-] / result valid flag
    bReorder : BOOL; // 补货标志（在手 ≤ 订货点）[-] / reorder flag
    iErrCode : INT; // 事件码 0=正常 1=日耗为负 2=提前期为负已归零 3=安全天数为负已归零 4=结果非有限 / event code
END_VAR
VAR
    rLeadUse : REAL; // 生效提前期 [d] / effective lead time
    rSafetyUse : REAL; // 生效安全天数 [d] / effective safety days
    rCoverDays : REAL; // 合计覆盖天数 [d] / total coverage days
    rRopRaw : REAL; // 未校验订货点 [件] / unchecked reorder point
    rShortRaw : REAL; // 未校验缺口量 [件] / unchecked shortage
END_VAR

    // —— 段 0：全路径预清 —— //
    rLeadUse := 0.0;
    rSafetyUse := 0.0;
    rCoverDays := 0.0;
    rRopRaw := 0.0;
    rShortRaw := 0.0;
    rRop := 0.0;
    rShortQty := 0.0;
    bValid := FALSE;
    bReorder := FALSE;
    iErrCode := 0;
    FC_DL_SpareReorderPoint := FALSE;
    // —— 段 1：日耗域闸（负消耗无物理意义） —— //
    IF rDailyUse < 0.0 THEN
        iErrCode := 1; // 日耗为负，订货点不可信 / negative daily use
        RETURN;
    END_IF;
    // —— 段 2：天数负值归零（配置错误宽容处理） —— //
    IF rLeadDays < 0.0 THEN
        rLeadUse := 0.0;
        iErrCode := 2; // 提前期为负已归零 / negative lead time clamped
    ELSE
        rLeadUse := rLeadDays;
    END_IF;
    IF rSafetyDays < 0.0 THEN
        rSafetyUse := 0.0;
        iErrCode := 3; // 安全天数为负已归零 / negative safety days clamped
    ELSE
        rSafetyUse := rSafetyDays;
    END_IF;
    // —— 段 3：量纲链 (件/d)×(d) = 件 —— //
    rCoverDays := rLeadUse + rSafetyUse; // 覆盖天数 [d] / coverage days
    rRopRaw := rDailyUse * rCoverDays; // 订货点 [件] / reorder point
    IF ABS(rRopRaw) > 1.0E15 THEN
        iErrCode := 4; // 结果非有限，强制归零 / non-finite result, forced to zero
        RETURN;
    END_IF;
    rRop := rRopRaw;
    // —— 段 4：缺口量 = MAX(0, 订货点-在手) 与补货判定 —— //
    rShortRaw := rRop - rOnHand; // 缺口 [件] / shortage
    IF rShortRaw < 0.0 THEN
        rShortQty := 0.0; // 库存充足，缺口为零 / enough stock
    ELSE
        rShortQty := rShortRaw;
    END_IF;
    bReorder := rOnHand <= rRop; // 补货标志 [-] / reorder flag
    bValid := TRUE;
    FC_DL_SpareReorderPoint := TRUE;
END_FUNCTION

(* ---- FC_DL_SprayFlowRateCalc.st ---- *)
(*
  Name: FC_DL_SprayFlowRateCalc
  Category: DL_Device
  Version: 1.0.0
  Round: R89 / 2026-11-25
  开源溯源：clean-room 自研（族 涂装喷涂线，ST 开源生态实测 0 命中，无外部代码引入）
  功能：喷枪流量与雾化压力匹配：按喷嘴孔径、供压、粘度算体积流量并按泵上限钳位，同时给出雾化压力建议值。
  边界条件：① 四入参全部过非有限闸，任一非有限返回哨兵 -1；
            ② 孔口流量用 Q = Cd·A·√(2ΔP/ρ)，Cd = 0.62、ρ = 1200 kg/m3 为涂料通用常量；
            ③ 粘度修正 kμ = 1/(1 + 0.3·√(ν/100))，ν 为运动粘度 [cSt]，量与基准同量纲故无量纲；
            ④ 雾化压力取供压的 85 % 并钳 0.5~6 bar（低压雾化枪工艺域），钳位只在量值上，不改有效性。
  量纲自证：m2 × √(Pa/(kg/m3)) = m2 × m/s = m3/s；m3/s × 1e6 = ml/s；×60 = ml/min。
*)
FUNCTION FC_DL_SprayFlowRateCalc : REAL
VAR_INPUT
    fNozzleDiaMm : REAL;        (* 喷嘴孔径 [mm] Nozzle orifice diameter [mm] *)
    fPressBar : REAL;           (* 供漆压力 [bar] Paint supply pressure [bar] *)
    fViscCst : REAL;            (* 运动粘度 [cSt] Kinematic viscosity [cSt] *)
    fFlowMaxMlmin : REAL;       (* 泵/枪流量上限 [ml/min] Flow ceiling [ml/min] *)
END_VAR
VAR_OUTPUT
    fFlowMlmin : REAL;          (* 计算流量（已钳位） [ml/min] Flow rate, clamped [ml/min] *)
    fAtomPressBar : REAL;       (* 雾化压力建议值 [bar] Recommended atomizing pressure [bar] *)
    xClamped : BOOL;            (* 流量已按上限钳位 [-] Flow clamped by ceiling *)
    xValid : BOOL;              (* 计算有效性标志 [-] Calculation valid flag *)
END_VAR
VAR CONSTANT
    DL_EPS : REAL := 1.0E-9;        (* 判据容差 [-] Criterion tolerance *)
    DL_CD : REAL := 0.62;           (* 孔口流量系数 [-] Orifice discharge coefficient *)
    DL_RHO : REAL := 1200.0;        (* 涂料密度（通用常量） [kg/m3] Paint density [kg/m3] *)
    DL_BAR_PA : REAL := 100000.0;   (* bar → Pa 换算 [Pa/bar] Bar to pascal *)
    DL_MM2_M2 : REAL := 1.0E6;      (* mm2 → m2 换算 [mm2/m2] Square millimetre to square metre *)
    DL_M3_ML : REAL := 1.0E6;       (* m3 → ml 换算 [ml/m3] Cubic metre to millilitre *)
    DL_SECMIN : REAL := 60.0;       (* 每秒 → 每分钟换算 [s/min] Second to minute *)
    DL_KVISC : REAL := 0.3;         (* 粘度修正系数 [-] Viscosity correction coefficient *)
    DL_VISC_REF : REAL := 100.0;    (* 粘度修正基准 [cSt] Viscosity reference [cSt] *)
    DL_ATOM_RATIO : REAL := 0.85;   (* 雾化压力/供压比 [-] Atomizing to supply ratio *)
    DL_ATOM_MIN : REAL := 0.5;      (* 雾化压力下限 [bar] Atomizing pressure floor [bar] *)
    DL_ATOM_MAX : REAL := 6.0;      (* 雾化压力上限 [bar] Atomizing pressure ceiling [bar] *)
    DL_PI_Q : REAL := 0.7853981633974483;  (* π/4（圆面积系数） [-] Quarter pi *)
    DL_DIA_MIN : REAL := 0.2;       (* 孔径下限 [mm] Diameter floor [mm] *)
    DL_DIA_MAX : REAL := 5.0;       (* 孔径上限 [mm] Diameter ceiling [mm] *)
    DL_P_MIN : REAL := 0.5;         (* 供压下限 [bar] Pressure floor [bar] *)
    DL_P_MAX : REAL := 10.0;        (* 供压上限 [bar] Pressure ceiling [bar] *)
    DL_V_MIN : REAL := 5.0;         (* 粘度下限 [cSt] Viscosity floor [cSt] *)
    DL_V_MAX : REAL := 2000.0;      (* 粘度上限 [cSt] Viscosity ceiling [cSt] *)
    DL_Q_MIN : REAL := 10.0;        (* 流量上限下限 [ml/min] Ceiling floor [ml/min] *)
    DL_Q_MAX : REAL := 5000.0;      (* 流量上限上限 [ml/min] Ceiling top [ml/min] *)
END_VAR
VAR
    fAreaM2 : REAL;     (* 孔口面积 [m2] Orifice area [m2] *)
    fDpPa : REAL;       (* 压差 [Pa] Differential pressure [Pa] *)
    fKvisc : REAL;      (* 粘度修正系数 [-] Viscosity correction factor *)
    fQm3s : REAL;       (* 体积流量 [m3/s] Volumetric flow [m3/s] *)
END_VAR
(* 出口预置：四出口统一预置（R256） *)
fFlowMlmin := 0.0; fAtomPressBar := 0.0; xClamped := FALSE; xValid := FALSE;
(* 非有限闸：NaN 自反判 + Inf 差值自减判，四入参全枚举 *)
IF (fNozzleDiaMm <> fNozzleDiaMm) OR ((fNozzleDiaMm - fNozzleDiaMm) <> 0.0)
   OR (fPressBar <> fPressBar) OR ((fPressBar - fPressBar) <> 0.0)
   OR (fViscCst <> fViscCst) OR ((fViscCst - fViscCst) <> 0.0)
   OR (fFlowMaxMlmin <> fFlowMaxMlmin) OR ((fFlowMaxMlmin - fFlowMaxMlmin) <> 0.0) THEN
    FC_DL_SprayFlowRateCalc := -1.0;        (* 哨兵 -1：入参非有限 / Sentinel -1, non-finite input *)
    RETURN;
END_IF
(* 组态域闸：孔径、供压、粘度、泵上限逐项定域 *)
IF (fNozzleDiaMm < DL_DIA_MIN) OR (fNozzleDiaMm > DL_DIA_MAX)
   OR (fPressBar < DL_P_MIN) OR (fPressBar > DL_P_MAX)
   OR (fViscCst < DL_V_MIN) OR (fViscCst > DL_V_MAX)
   OR (fFlowMaxMlmin < DL_Q_MIN) OR (fFlowMaxMlmin > DL_Q_MAX) THEN
    FC_DL_SprayFlowRateCalc := -1.0;        (* 哨兵 -1：组态非法 / Sentinel -1, bad configuration *)
    RETURN;
END_IF
(* 孔口面积：π/4·d² [mm2] ÷ 1e6 = m2 *)
fAreaM2 := (DL_PI_Q * fNozzleDiaMm * fNozzleDiaMm) / DL_MM2_M2;
(* 压差：bar × 1e5 = Pa *)
fDpPa := fPressBar * DL_BAR_PA;
(* 粘度修正：ν/100 无量纲，开方后按 0.3 权重并入分母，恒在 (0, 1] 区间 *)
fKvisc := 1.0 / (1.0 + DL_KVISC * SQRT(fViscCst / DL_VISC_REF));
(* 孔口流量：m2 × √(Pa/(kg/m3)) = m2 × m/s = m3/s *)
fQm3s := DL_CD * fAreaM2 * SQRT((2.0 * fDpPa) / DL_RHO) * fKvisc;
(* 单位换算：m3/s → ml/min *)
fFlowMlmin := fQm3s * DL_M3_ML * DL_SECMIN;
(* 泵上限钳位：置钳位标志，有效性不变（事实未伪造） *)
IF fFlowMlmin > fFlowMaxMlmin THEN
    fFlowMlmin := fFlowMaxMlmin;
    xClamped := TRUE;
END_IF
(* 雾化压力：供压 85 %，钳 0.5~6 bar *)
fAtomPressBar := fPressBar * DL_ATOM_RATIO;
IF fAtomPressBar < DL_ATOM_MIN THEN
    fAtomPressBar := DL_ATOM_MIN;
ELSIF fAtomPressBar > DL_ATOM_MAX THEN
    fAtomPressBar := DL_ATOM_MAX;
END_IF
xValid := TRUE;                             (* 链路有效 / Chain valid *)
FC_DL_SprayFlowRateCalc := fFlowMlmin;
END_FUNCTION

(* ---- FC_DL_SpreaderTwistLockChk.st ---- *)
(*
 * FC_DL_SpreaderTwistLockChk | C2 | DL_Device
 * 功能：吊具四角旋锁的到位互锁判定（全锁 / 全开 / 未知 / 故障）       单位：nLockState [枚举码 0/1/2/3]、nFaultCode [INT]
 * 工况边界：仅适用于四角独立旋锁（每角一锁到位 + 一开到位双反馈）；单角双 ON、混合状态、计数越界一律判故障 9201 并置 xFault；本件为纯函数，超时由调用方 FB 计时
 * 代数值回代：四锁位全 ON 且四开位全 OFF → nLockState=1、xLockedOk=TRUE；四锁位全 OFF 且四开位全 ON → nLockState=2、xUnlockedOk=TRUE（与 spec 判定表一致）
 * 开源溯源：clean-room 自研，未复制任何第三方代码（无外部来源）
 *)
FUNCTION FC_DL_SpreaderTwistLockChk : BOOL
VAR_INPUT
    xLockFL   : BOOL;                // 左前锁到位 | front-left locked
    xLockFR   : BOOL;                // 右前锁到位 | front-right locked
    xLockRL   : BOOL;                // 左后锁到位 | rear-left locked
    xLockRR   : BOOL;                // 右后锁到位 | rear-right locked
    xUnlockFL : BOOL;                // 左前开到位 | front-left unlocked
    xUnlockFR : BOOL;                // 右前开到位 | front-right unlocked
    xUnlockRL : BOOL;                // 左后开到位 | rear-left unlocked
    xUnlockRR : BOOL;                // 右后开到位 | rear-right unlocked
END_VAR
VAR_OUTPUT
    nLockState : INT;                // 0=未知 / 1=全锁 / 2=全开 / 3=故障 | 0 unknown, 1 all locked, 2 all unlocked, 3 fault
    xLockedOk  : BOOL;               // 允许起吊（四角全锁）| lifting permitted, all four locked
    xUnlockedOk: BOOL;               // 允许脱箱（四角全开）| releasing permitted, all four unlocked
    xFault     : BOOL;               // 故障标志 | fault flag
    nFaultCode : INT;                // 故障码 0=无 / 9201=旋锁状态非法 | fault code 0=none, 9201=illegal twist lock state
    xValid     : BOOL;               // 判定结果可用（全锁或全开）| the verdict is usable, all locked or all unlocked
END_VAR
VAR
    nLockOn   : INT;                 // 锁到位计数 | count of locked positions
    nUnlockOn : INT;                 // 开到位计数 | count of unlocked positions
END_VAR

// 段1｜计数：分别统计锁到位与开到位（同角双 ON 会体现在计数总和中）
nLockOn := 0;
nUnlockOn := 0;
IF xLockFL THEN
    nLockOn := nLockOn + 1;
END_IF
IF xLockFR THEN
    nLockOn := nLockOn + 1;
END_IF
IF xLockRL THEN
    nLockOn := nLockOn + 1;
END_IF
IF xLockRR THEN
    nLockOn := nLockOn + 1;
END_IF
IF xUnlockFL THEN
    nUnlockOn := nUnlockOn + 1;
END_IF
IF xUnlockFR THEN
    nUnlockOn := nUnlockOn + 1;
END_IF
IF xUnlockRL THEN
    nUnlockOn := nUnlockOn + 1;
END_IF
IF xUnlockRR THEN
    nUnlockOn := nUnlockOn + 1;
END_IF

// 段2｜状态判定（出口先取安全侧：不允许起吊也不允许脱箱）
xLockedOk := FALSE;
xUnlockedOk := FALSE;
xFault := FALSE;
nFaultCode := 0;
IF (nLockOn = 4) AND (nUnlockOn = 0) THEN
    nLockState := 1;                 // 全锁：四锁位 ON + 四开位 OFF | all locked
    xLockedOk := TRUE;
ELSIF (nLockOn = 0) AND (nUnlockOn = 4) THEN
    nLockState := 2;                 // 全开：四开位 ON + 四锁位 OFF | all unlocked
    xUnlockedOk := TRUE;
ELSIF (nLockOn = 0) AND (nUnlockOn = 0) THEN
    nLockState := 0;                 // 未知：无任何到位反馈 | unknown, no feedback at all
ELSIF (nLockOn + nUnlockOn) > 4 THEN
    nLockState := 3;                 // 故障：同角双 ON 或计数越界 | fault, both bits of one corner are on
    xFault := TRUE;
    nFaultCode := 9201;
ELSE
    nLockState := 3;                 // 故障：混合状态（部分锁部分开）| fault, mixed state
    xFault := TRUE;
    nFaultCode := 9201;
END_IF

// 段3｜出口：只有全锁或全开才认为判定可用
xValid := xLockedOk OR xUnlockedOk;
FC_DL_SpreaderTwistLockChk := xValid;
END_FUNCTION

(* ---- FC_DL_StrainBridgeExcitationComp.st ---- *)
(* ===========================================================================
   组件名   : FC_DL_StrainBridgeExcitationComp
   分类     : DL_Device / 桥压激励补偿
   一句话   : 按实测激励电压与额定值之比归一化桥路输出，消除激励波动引起的比例误差
   复杂度   : 1        版本 : v1.0.0        日期 : 2026-11-24
   开源溯源 : 无（clean-room 自研，未借鉴任何开源实现）
   输入契约 : fRawValue 原始读数（已换算值）；fExcMeasV 实测激励电压 [V]
              fExcRatedV 额定激励电压 [V]；fRatioMin/fRatioMax 比例合理区间
   输出契约 : 返回值 = 归一化后读数；fRatio 归一化比例（额定/实测）
              xValid 输入有效（比例须落在合理区间内）
   修改记录 : v1.0.0 2026-11-24 初版
   =========================================================================== *)

FUNCTION FC_DL_StrainBridgeExcitationComp : REAL
VAR_INPUT
    fRawValue : REAL;                  // 原始读数 | raw reading
    fExcMeasV : REAL := 5.0;           // 实测激励电压 [V] | measured excitation [V]
    fExcRatedV : REAL := 5.0;          // 额定激励电压 [V] | rated excitation [V]
    fRatioMin : REAL := 0.5;           // 比例下限 | ratio lower bound
    fRatioMax : REAL := 2.0;           // 比例上限 | ratio upper bound
END_VAR
VAR_OUTPUT
    fRatio : REAL;                     // 归一化比例 | normalization ratio
    xValid : BOOL;                     // 输入有效标志 | inputs valid flag
END_VAR
VAR
    _fR : REAL;                        // 比例工作值 | ratio working value
    _fOut : REAL;                      // 归一化结果 | normalized result
END_VAR

// ---- 输出预置 ----
fRatio := 1.0;
xValid := FALSE;
FC_DL_StrainBridgeExcitationComp := 0.0;

// ---- 非有限值拦截 ----
IF (fRawValue <> fRawValue) OR ((fRawValue - fRawValue) <> (fRawValue - fRawValue)) THEN
    RETURN;
END_IF
IF (fExcMeasV <> fExcMeasV) OR ((fExcMeasV - fExcMeasV) <> (fExcMeasV - fExcMeasV)) THEN
    RETURN;
END_IF
IF (fExcRatedV <> fExcRatedV) OR ((fExcRatedV - fExcRatedV) <> (fExcRatedV - fExcRatedV)) THEN
    RETURN;
END_IF

// ---- 防除零：实测与额定激励都必须显著非零 ----
IF (ABS(fExcMeasV) < 0.000000001) OR (ABS(fExcRatedV) < 0.000000001) THEN
    RETURN;
END_IF

// ---- 比例 = 额定 / 实测 ----
_fR := fExcRatedV / fExcMeasV;                     // 分母已守卫
fRatio := _fR;

// ---- 合理性区间守卫：比例越界说明激励异常，宁判无效也不外推 ----
IF (fRatioMin <= 0.0) OR (fRatioMax <= fRatioMin) THEN
    RETURN;
END_IF
IF (_fR < fRatioMin) OR (_fR > fRatioMax) THEN
    RETURN;
END_IF

_fOut := fRawValue * _fR;
xValid := TRUE;
FC_DL_StrainBridgeExcitationComp := _fOut;
END_FUNCTION

(* ---- FC_DL_StrainBridgeMillivolt.st ---- *)
(* ===========================================================================
   组件名   : FC_DL_StrainBridgeMillivolt
   分类     : DL_Device / 应变桥信号换算
   一句话   : 由激励电压与实测差分电压算桥路输出 mV/V 与等效微应变
   复杂度   : 1        版本 : v1.0.0        日期 : 2026-11-24
   开源溯源 : 无（clean-room 自研，未借鉴任何开源实现）
   输入契约 : fExcitationV 桥路激励电压 [V]；fDiffV 实测差分电压 [mV]
              fGaugeFactor 应变片灵敏系数（典型 2.0）
   输出契约 : 返回值 = 桥路输出 [mV/V]；fMvPerV 同返回值（显式输出）
              fMicroStrain 等效微应变 [µε]（= mV/V × 1000 / GF）；xValid 输入有效
   修改记录 : v1.0.0 2026-11-24 初版
   =========================================================================== *)

FUNCTION FC_DL_StrainBridgeMillivolt : REAL
VAR_INPUT
    fExcitationV : REAL := 5.0;        // 桥路激励电压 [V] | bridge excitation [V]
    fDiffV : REAL;                     // 实测差分电压 [mV] | measured differential [mV]
    fGaugeFactor : REAL := 2.0;        // 应变片灵敏系数 | gauge factor
END_VAR
VAR_OUTPUT
    fMvPerV : REAL;                    // 桥路输出 [mV/V] | bridge output [mV/V]
    fMicroStrain : REAL;               // 等效微应变 [µε] | equivalent micro strain [µε]
    xValid : BOOL;                     // 输入有效标志 | inputs valid flag
END_VAR
VAR
    _fRatio : REAL;                    // 差分/激励 比值 | differential over excitation
END_VAR

// ---- 输出预置 ----
fMvPerV := 0.0;
fMicroStrain := 0.0;
xValid := FALSE;
FC_DL_StrainBridgeMillivolt := 0.0;

// ---- 非有限值拦截 ----
IF (fExcitationV <> fExcitationV) OR ((fExcitationV - fExcitationV) <> (fExcitationV - fExcitationV)) THEN
    RETURN;
END_IF
IF (fDiffV <> fDiffV) OR ((fDiffV - fDiffV) <> (fDiffV - fDiffV)) THEN
    RETURN;
END_IF
IF (fGaugeFactor <> fGaugeFactor) OR ((fGaugeFactor - fGaugeFactor) <> (fGaugeFactor - fGaugeFactor)) THEN
    RETURN;
END_IF

// ---- 防除零：激励电压与灵敏系数必须显著非零 ----
IF (ABS(fExcitationV) < 0.000000001) OR (ABS(fGaugeFactor) < 0.000000001) THEN
    RETURN;
END_IF

// ---- mV/V = 差分电压 [mV] / 激励电压 [V] ----
_fRatio := fDiffV / fExcitationV;                  // 分母已守卫
fMvPerV := _fRatio;

// ---- 微应变 = (mV/V) × 1000 / GF，全桥条件下 GF=2 时 1 mV/V ≈ 500 µε ----
fMicroStrain := _fRatio * 1000.0 / fGaugeFactor;   // 分母已守卫

xValid := TRUE;
FC_DL_StrainBridgeMillivolt := _fRatio;
END_FUNCTION

(* ---- FC_DL_StrainBridgeNonlinCorr.st ---- *)
(* ===========================================================================
   组件名   : FC_DL_StrainBridgeNonlinCorr
   分类     : DL_Device / 桥路非线性修正
   一句话   : 用三次多项式修正大应变下桥路输出的非线性误差，保留原始符号
   复杂度   : 2        版本 : v1.0.0        日期 : 2026-11-24
   开源溯源 : 无（clean-room 自研，未借鉴任何开源实现）
   输入契约 : fRawStrain 原始应变 [µε]；fK2 二次项系数 [1/µε]；fK3 三次项系数 [1/µε²]
   输出契约 : 返回值 = 修正后应变 [µε]；fCorrTerm 修正量 [µε]；xValid 输入有效
   算法说明 : ε_corr = ε_raw + K2·ε_raw² + K3·ε_raw³；二次项破坏奇对称性，故系数须由标定给定，
              未标定时置 0 即为旁路；输入超过 ±1e6 µε 视为超量程而判无效
   修改记录 : v1.0.0 2026-11-24 初版
   =========================================================================== *)

FUNCTION FC_DL_StrainBridgeNonlinCorr : REAL
VAR_INPUT
    fRawStrain : REAL;                 // 原始应变 [µε] | raw strain [µε]
    fK2 : REAL := 0.0;                 // 二次项系数 [1/µε] | quadratic coefficient [1/µε]
    fK3 : REAL := 0.0;                 // 三次项系数 [1/µε²] | cubic coefficient [1/µε^2]
    fRangeLimit : REAL := 1000000.0;   // 量程上限 [µε] | range limit [µε]
END_VAR
VAR_OUTPUT
    fCorrTerm : REAL;                  // 修正量 [µε] | correction term [µε]
    xValid : BOOL;                     // 输入有效标志 | inputs valid flag
END_VAR
VAR
    _fSq : REAL;                       // 应变平方 [(µε)²] | squared strain
    _fCub : REAL;                      // 应变立方 [(µε)³] | cubed strain
    _fOut : REAL;                      // 修正结果 [µε] | corrected result [µε]
END_VAR

// ---- 输出预置 ----
fCorrTerm := 0.0;
xValid := FALSE;
FC_DL_StrainBridgeNonlinCorr := 0.0;

// ---- 非有限值拦截 ----
IF (fRawStrain <> fRawStrain) OR ((fRawStrain - fRawStrain) <> (fRawStrain - fRawStrain)) THEN
    RETURN;
END_IF
IF (fK2 <> fK2) OR ((fK2 - fK2) <> (fK2 - fK2)) THEN
    RETURN;
END_IF
IF (fK3 <> fK3) OR ((fK3 - fK3) <> (fK3 - fK3)) THEN
    RETURN;
END_IF

// ---- 量程守卫：上限非正或超量程一律判无效，避免三次项数值爆炸 ----
IF (fRangeLimit <= 0.0) THEN
    RETURN;
END_IF
IF ABS(fRawStrain) > fRangeLimit THEN
    RETURN;
END_IF

// ---- 多项式修正：先算平方与立方再合成，避免重复乘法产生不同舍入路径 ----
_fSq := fRawStrain * fRawStrain;
_fCub := _fSq * fRawStrain;
fCorrTerm := fK2 * _fSq + fK3 * _fCub;
_fOut := fRawStrain + fCorrTerm;

// ---- 结果二次守卫：修正后仍须在量程内，否则判无效 ----
IF ABS(_fOut) > (fRangeLimit * 2.0) THEN
    xValid := FALSE;
    RETURN;
END_IF

xValid := TRUE;
FC_DL_StrainBridgeNonlinCorr := _fOut;
END_FUNCTION

(* ---- FC_DL_StrainCreepComp.st ---- *)
(* ===========================================================================
   组件名   : FC_DL_StrainCreepComp
   分类     : DL_Device / 应变蠕变补偿
   一句话   : 按载荷保持时间与蠕变系数用指数饱和模型修正读数漂移
   复杂度   : 2        版本 : v1.0.0        日期 : 2026-11-24
   开源溯源 : 无（clean-room 自研，未借鉴任何开源实现）
   输入契约 : fRawStrain 原始应变 [µε]；fHoldSec 载荷保持时间 [s]
              fCreepK 蠕变系数（0..0.1，无量纲） | creep coefficient
              fTauSec 蠕变时间常数 [s]
   输出契约 : 返回值 = 蠕变修正后应变 [µε]；fCreepTerm 蠕变量 [µε]
              fCreepFrac 蠕变完成度 0..1；xValid 输入有效
   修改记录 : v1.0.0 2026-11-24 初版
   =========================================================================== *)

FUNCTION FC_DL_StrainCreepComp : REAL
VAR_INPUT
    fRawStrain : REAL;                 // 原始应变 [µε] | raw strain [µε]
    fHoldSec : REAL := 0.0;            // 载荷保持时间 [s] | load hold time [s]
    fCreepK : REAL := 0.01;            // 蠕变系数 0..0.1 | creep coefficient 0..0.1
    fTauSec : REAL := 60.0;            // 蠕变时间常数 [s] | creep time constant [s]
END_VAR
VAR_OUTPUT
    fCreepTerm : REAL;                 // 蠕变量 [µε] | creep amount [µε]
    fCreepFrac : REAL;                 // 蠕变完成度 0..1 | creep completion 0..1
    xValid : BOOL;                     // 输入有效标志 | inputs valid flag
END_VAR
VAR
    _fRatio : REAL;                    // 保持时间/时间常数 | hold over tau
    _fFrac : REAL;                     // 蠕变完成度 | creep completion
    _fOut : REAL;                      // 修正结果 [µε] | corrected result [µε]
END_VAR

// ---- 输出预置 ----
fCreepTerm := 0.0;
fCreepFrac := 0.0;
xValid := FALSE;
FC_DL_StrainCreepComp := 0.0;

// ---- 非有限值拦截 ----
IF (fRawStrain <> fRawStrain) OR ((fRawStrain - fRawStrain) <> (fRawStrain - fRawStrain)) THEN
    RETURN;
END_IF
IF (fHoldSec <> fHoldSec) OR ((fHoldSec - fHoldSec) <> (fHoldSec - fHoldSec)) THEN
    RETURN;
END_IF
IF (fCreepK <> fCreepK) OR ((fCreepK - fCreepK) <> (fCreepK - fCreepK)) THEN
    RETURN;
END_IF
IF (fTauSec <> fTauSec) OR ((fTauSec - fTauSec) <> (fTauSec - fTauSec)) THEN
    RETURN;
END_IF

// ---- 防除零与参数守卫：时间常数必须为正，蠕变系数限于 0..0.1 ----
IF (fTauSec < 0.000001) OR (fCreepK < 0.0) OR (fCreepK > 0.1) OR (fHoldSec < 0.0) THEN
    RETURN;
END_IF

// ---- 指数饱和模型：完成度 = 1 − exp(−t/τ)，比值上限 50 防下溢 ----
_fRatio := fHoldSec / fTauSec;                     // 分母已守卫
IF _fRatio > 50.0 THEN
    _fRatio := 50.0;
END_IF
_fFrac := 1.0 - EXP(-_fRatio);
fCreepFrac := _fFrac;

// ---- 蠕变量按原始读数比例给出，再从读数中扣除 ----
fCreepTerm := fRawStrain * fCreepK * _fFrac;
_fOut := fRawStrain - fCreepTerm;

xValid := TRUE;
FC_DL_StrainCreepComp := _fOut;
END_FUNCTION

(* ---- FC_DL_StrainGaugeTempComp.st ---- *)
(* ===========================================================================
   组件名   : FC_DL_StrainGaugeTempComp
   分类     : DL_Device / 应变片温度补偿
   一句话   : 按敏感栅与补偿片温差、灵敏系数温度系数对读数做灵敏度与零点双重修正
   复杂度   : 2        版本 : v1.0.0        日期 : 2026-11-24
   开源溯源 : 无（clean-room 自研，未借鉴任何开源实现）
   输入契约 : fRawStrain 原始读数 [µε]；fTempSens 敏感栅温度 [°C]；fTempComp 补偿片温度 [°C]
              fRefTemp 参考温度 [°C]；fTkSens 灵敏系数温度系数 [1/°C]
              fTkZero 零点温度漂移系数 [µε/°C]
   输出契约 : 返回值 = 修正后应变 [µε]；fSensFactor 灵敏度修正因子
              fZeroShift 零点漂移修正量 [µε]；fDeltaTSens 敏感栅温差 [°C]；xValid 输入有效
   修改记录 : v1.0.0 2026-11-24 初版
   =========================================================================== *)

FUNCTION FC_DL_StrainGaugeTempComp : REAL
VAR_INPUT
    fRawStrain : REAL;                 // 原始读数 [µε] | raw strain reading [µε]
    fTempSens : REAL := 25.0;          // 敏感栅温度 [°C] | sensing grid temperature [°C]
    fTempComp : REAL := 25.0;          // 补偿片温度 [°C] | compensation grid temperature [°C]
    fRefTemp : REAL := 20.0;           // 参考温度 [°C] | reference temperature [°C]
    fTkSens : REAL := 0.0002;          // 灵敏系数温度系数 [1/°C] | tc of gauge factor [1/°C]
    fTkZero : REAL := 1.0;             // 零点温度漂移系数 [µε/°C] | zero tc [µε/°C]
END_VAR
VAR_OUTPUT
    fSensFactor : REAL;                // 灵敏度修正因子 | sensitivity correction factor
    fZeroShift : REAL;                 // 零点漂移修正量 [µε] | zero shift correction [µε]
    fDeltaTSens : REAL;                // 敏感栅温差 [°C] | sensing grid temp delta [°C]
    xValid : BOOL;                     // 输入有效标志 | inputs valid flag
END_VAR
VAR
    _fOut : REAL;                      // 修正结果 [µε] | corrected result [µε]
END_VAR

// ---- 输出预置 ----
fSensFactor := 1.0;
fZeroShift := 0.0;
fDeltaTSens := 0.0;
xValid := FALSE;
FC_DL_StrainGaugeTempComp := 0.0;

// ---- 非有限值拦截 ----
IF (fRawStrain <> fRawStrain) OR ((fRawStrain - fRawStrain) <> (fRawStrain - fRawStrain)) THEN
    RETURN;
END_IF
IF (fTempSens <> fTempSens) OR ((fTempSens - fTempSens) <> (fTempSens - fTempSens)) THEN
    RETURN;
END_IF
IF (fTempComp <> fTempComp) OR ((fTempComp - fTempComp) <> (fTempComp - fTempComp)) THEN
    RETURN;
END_IF
IF (fRefTemp <> fRefTemp) OR ((fRefTemp - fRefTemp) <> (fRefTemp - fRefTemp)) THEN
    RETURN;
END_IF

// ---- 温差计算：敏感栅温差用于灵敏度修正，补偿片温差用于零点修正 ----
fDeltaTSens := fTempSens - fRefTemp;
fSensFactor := 1.0 + fTkSens * fDeltaTSens;
fZeroShift := fTkZero * (fTempComp - fRefTemp);

// ---- 防除零：灵敏度因子必须显著非零 ----
IF ABS(fSensFactor) < 0.000000001 THEN
    RETURN;
END_IF

// ---- 先除灵敏度因子消去灵敏度温漂，再扣零点温漂 ----
_fOut := fRawStrain / fSensFactor - fZeroShift;     // 分母已守卫

xValid := TRUE;
FC_DL_StrainGaugeTempComp := _fOut;
END_FUNCTION

(* ---- FC_DL_StrainMultiPointCalib.st ---- *)
(* ===========================================================================
   组件名   : FC_DL_StrainMultiPointCalib
   分类     : DL_Device / 应变多点标定插值
   一句话   : 按标定点表分段线性插值反算工程量，段号钳位并对表外输入做平段外推
   复杂度   : 2        版本 : v1.0.0        日期 : 2026-11-24
   开源溯源 : 无（clean-room 自研，未借鉴任何开源实现）
   输入契约 : fRaw 原始读数 [µε]；afRawPT 标定原始值表 [1..8]；afEngPT 标定工程量表 [1..8]
              iCount 有效点数 2..8（自动钳位）
   输出契约 : 返回值 = 工程量；iSeg 命中的段号（1..iCount−1）；fRawClamped 钳位后原始值
              xValid 表数据有效（升序且有限）
   修改记录 : v1.0.0 2026-11-24 初版
   =========================================================================== *)

FUNCTION FC_DL_StrainMultiPointCalib : REAL
VAR_INPUT
    fRaw : REAL;                       // 原始读数 [µε] | raw reading [µε]
    afRawPT : ARRAY[1..8] OF REAL;     // 标定原始值表 | calibration raw points
    afEngPT : ARRAY[1..8] OF REAL;     // 标定工程量表 | calibration engineering points
    iCount : INT := 8;                 // 有效点数 2..8 | valid point count 2..8
END_VAR
VAR_OUTPUT
    iSeg : INT;                        // 命中段号 | hit segment index
    fRawClamped : REAL;                // 钳位后原始值 [µε] | clamped raw value [µε]
    xValid : BOOL;                     // 输入有效标志 | inputs valid flag
END_VAR
VAR
    _iN : INT;                         // 钳位后点数 | clamped point count
    _i : INT;                          // 循环下标 | loop index
    _fDen : REAL;                      // 段宽 | segment width
    _fSlope : REAL;                    // 段斜率 | segment slope
    _fOut : REAL;                      // 插值结果 | interpolation result
    _xMono : BOOL;                     // 表单调升序标志 | monotonic ascending flag
END_VAR

// ---- 输出预置 ----
iSeg := 1;
fRawClamped := 0.0;
xValid := FALSE;
FC_DL_StrainMultiPointCalib := 0.0;

// ---- 非有限值拦截 ----
IF (fRaw <> fRaw) OR ((fRaw - fRaw) <> (fRaw - fRaw)) THEN
    RETURN;
END_IF

// ---- 点数钳位：至少 2 点，最多 8 点 ----
_iN := iCount;
IF _iN < 2 THEN
    _iN := 2;
ELSIF _iN > 8 THEN
    _iN := 8;
END_IF

// ---- 表数据校验：全部有限且原始值严格升序（插值前提） ----
_xMono := TRUE;
_i := 1;
WHILE _i <= _iN DO
    IF (afRawPT[_i] <> afRawPT[_i]) OR ((afRawPT[_i] - afRawPT[_i]) <> (afRawPT[_i] - afRawPT[_i])) THEN
        _xMono := FALSE;
    END_IF
    IF (afEngPT[_i] <> afEngPT[_i]) OR ((afEngPT[_i] - afEngPT[_i]) <> (afEngPT[_i] - afEngPT[_i])) THEN
        _xMono := FALSE;
    END_IF
    IF _i >= 2 THEN
        IF (afRawPT[_i] - afRawPT[_i - 1]) <= 0.000000001 THEN
            _xMono := FALSE;                       // 非严格升序即判表非法
        END_IF
    END_IF
    _i := _i + 1;
END_WHILE
IF NOT _xMono THEN
    RETURN;
END_IF

// ---- 输入钳位到标定区间：表外输入按平段外推，不外插 ----
_fOut := fRaw;
IF fRaw < afRawPT[1] THEN
    _fOut := afRawPT[1];
ELSIF fRaw > afRawPT[_iN] THEN
    _fOut := afRawPT[_iN];
END_IF
fRawClamped := _fOut;

// ---- 定位命中段：段号限制在 1.._iN−1，防数组越界 ----
iSeg := 1;
_i := 1;
WHILE _i <= (_iN - 1) DO
    IF (_fOut >= afRawPT[_i]) AND (_fOut <= afRawPT[_i + 1]) THEN
        iSeg := _i;                                // 命中区间 [i, i+1]
    END_IF
    _i := _i + 1;
END_WHILE
IF iSeg < 1 THEN
    iSeg := 1;
ELSIF iSeg > (_iN - 1) THEN
    iSeg := _iN - 1;                               // 下标钳位
END_IF

// ---- 分段线性插值 ----
_fDen := afRawPT[iSeg + 1] - afRawPT[iSeg];
IF ABS(_fDen) < 0.000000001 THEN
    _fSlope := 0.0;                                // 段宽为零则退化为平段，避免除零
ELSE
    _fSlope := (afEngPT[iSeg + 1] - afEngPT[iSeg]) / _fDen;   // 分母已守卫
END_IF
_fOut := afEngPT[iSeg] + (_fOut - afRawPT[iSeg]) * _fSlope;

xValid := TRUE;
FC_DL_StrainMultiPointCalib := _fOut;
END_FUNCTION

(* ---- FC_DL_StrainRosettePrincipal.st ---- *)
(* ===========================================================================
   组件名   : FC_DL_StrainRosettePrincipal
   分类     : DL_Device / 应变花主应变
   一句话   : 由 0°/45°/90° 三向应变算主应变、主方向角与最大剪应变
   复杂度   : 3        版本 : v1.0.0        日期 : 2026-11-24
   开源溯源 : 无（clean-room 自研，未借鉴任何开源实现）
   输入契约 : fEpsA 0° 应变 [µε]；fEpsB 45° 应变 [µε]；fEpsC 90° 应变 [µε]
   输出契约 : 返回值 = 第一主应变 ε1 [µε]
              fEps2 第二主应变 [µε]；fAngRad 主方向角 [rad]（−π/2, π/2]
              fShearMax 最大剪应变 [µε]；fCenter 应变圆心 [µε]；xValid 输入有效
   算法说明 : 令 C=(a+c)/2、A=(a−c)/2、B=(2b−a−c)/2，则 ε(θ)=C+A·cos2θ+B·sin2θ
              ε1,2 = C ± √(A²+B²)，2θp = atan2(B, A)，θp = 0.5·atan2(B, A)
   修改记录 : v1.0.0 2026-11-24 初版
   =========================================================================== *)

FUNCTION FC_DL_StrainRosettePrincipal : REAL
VAR_INPUT
    fEpsA : REAL;                      // 0° 向应变 [µε] | 0 deg strain [µε]
    fEpsB : REAL;                      // 45° 向应变 [µε] | 45 deg strain [µε]
    fEpsC : REAL;                      // 90° 向应变 [µε] | 90 deg strain [µε]
END_VAR
VAR_OUTPUT
    fEps2 : REAL;                      // 第二主应变 [µε] | second principal strain [µε]
    fAngRad : REAL;                    // 主方向角 [rad] | principal direction [rad]
    fShearMax : REAL;                  // 最大剪应变 [µε] | maximum shear strain [µε]
    fCenter : REAL;                    // 应变圆心 [µε] | strain circle center [µε]
    xValid : BOOL;                     // 输入有效标志 | inputs valid flag
END_VAR
VAR
    _fC : REAL;                        // 圆心 (a+c)/2 [µε] | center [µε]
    _fA : REAL;                        // 余弦分量 (a−c)/2 [µε] | cosine component [µε]
    _fB : REAL;                        // 正弦分量 (2b−a−c)/2 [µε] | sine component [µε]
    _fR : REAL;                        // 半径（最大剪应变） [µε] | radius [µε]
    _fAng2 : REAL;                     // 二倍主方向角 [rad] | twice principal angle [rad]
    _fAng : REAL;                      // 主方向角 [rad] | principal angle [rad]
END_VAR

// ---- 输出预置 ----
fEps2 := 0.0;
fAngRad := 0.0;
fShearMax := 0.0;
fCenter := 0.0;
xValid := FALSE;
FC_DL_StrainRosettePrincipal := 0.0;

// ---- 非有限值拦截 ----
IF (fEpsA <> fEpsA) OR ((fEpsA - fEpsA) <> (fEpsA - fEpsA)) THEN
    RETURN;
END_IF
IF (fEpsB <> fEpsB) OR ((fEpsB - fEpsB) <> (fEpsB - fEpsB)) THEN
    RETURN;
END_IF
IF (fEpsC <> fEpsC) OR ((fEpsC - fEpsC) <> (fEpsC - fEpsC)) THEN
    RETURN;
END_IF

// ---- 应变圆三要素 ----
_fC := (fEpsA + fEpsC) * 0.5;
_fA := (fEpsA - fEpsC) * 0.5;
_fB := (2.0 * fEpsB - fEpsA - fEpsC) * 0.5;
fCenter := _fC;
_fR := SQRT(_fA * _fA + _fB * _fB);                // 平方和非负，SQRT 安全
fShearMax := _fR;

// ---- 主应变 ----
FC_DL_StrainRosettePrincipal := _fC + _fR;
fEps2 := _fC - _fR;

// ---- 手工 atan2：避免依赖非标准 ATAN2，先判分母再补象限 ----
_fAng2 := 0.0;
IF ABS(_fA) < 0.000000001 THEN
    IF _fB > 0.0 THEN
        _fAng2 := 1.570796327;                     // 分母近零且 B>0 → +π/2
    ELSIF _fB < 0.0 THEN
        _fAng2 := -1.570796327;                    // 分母近零且 B<0 → −π/2
    END_IF
ELSE
    _fAng2 := ATAN(_fB / _fA);                     // 分母已守卫
    IF _fA < 0.0 THEN
        IF _fB >= 0.0 THEN
            _fAng2 := _fAng2 + 3.141592654;        // 第二象限补偿
        ELSE
            _fAng2 := _fAng2 - 3.141592654;        // 第三象限补偿
        END_IF
    END_IF
END_IF

// ---- 主方向角：除以 2 并归一化到 (−π/2, π/2] ----
_fAng := _fAng2 * 0.5;
IF _fAng > 1.570796327 THEN
    _fAng := _fAng - 3.141592654;
ELSIF _fAng <= -1.570796327 THEN
    _fAng := _fAng + 3.141592654;
END_IF
fAngRad := _fAng;

xValid := TRUE;
END_FUNCTION

(* ---- FC_DL_StrandTensionAtWinderCalc.st ---- *)
// FC_DL_StrandTensionAtWinderCalc v1.0.0
// 开源溯源：clean-room 自研（族 DL_Device，ST 生态实测 0 命中，无外部代码引入）
(*
  功能: 有效总张力 = 总张力 − 导纱摩擦损失 + 线密度·加速度 [N]（惯性力项 m'·a），
        单束张力 = 有效总张力/丝束根数，×100 换算为 cN。
  邻件/码位: 与 FC_DL_SizeApplicatorPickupCalc 同属拉丝后端件（力学面 vs 化学面）；
             16#0002_9226 = 非有限、根数 < 1、摩擦/线密度为负或有效总张力非正拒收。
*)
FUNCTION FC_DL_StrandTensionAtWinderCalc : REAL
VAR_INPUT
    fTotalTension : REAL := 60.0;  // 总张力 [N]，域 > 0 / Total tension [N]
    iStrandCount  : INT := 400;     // 丝束根数，域 >= 1 [根] / Strand count
    fFrictionDrop : REAL := 2.0;    // 导纱摩擦损失 [N]，域 >= 0 / Guide friction drop [N]
    fAccel        : REAL := 0.5;    // 卷绕加速度 [m/s²] / Winding acceleration [m/s^2]
    fMassPerLen   : REAL := 0.02;   // 线密度 [kg/m]，域 >= 0 / Linear mass density [kg/m]
END_VAR
VAR_OUTPUT
    fTensionPerStrand : REAL;       // 单束张力 [cN] / Tension per strand [cN]
    bValid            : BOOL;       // 结果有效回执 [-] / Result validity receipt
    uErrorId          : UDINT;      // 事件码，0 = 无事件 / Event code
END_VAR
VAR
    fEffective : REAL := 0.0;       // 有效总张力 [N] / Effective total tension [N]
END_VAR
// 段 0：全路径出口安全缺省 / Safe defaults on all outlets
fTensionPerStrand := 0.0;           // 单束张力缺省零 / Per-strand default zero
bValid := FALSE;                    // 有效回执预清 / Validity preset clear
uErrorId := 16#0000;                // 事件码预清 / Event code preset clear
FC_DL_StrandTensionAtWinderCalc := 0.0;     // 返回值缺省零（镜像单束张力）/ Return default zero
// 段 1：非有限闸（四实数入参；整数入参天然有限）/ Non-finite gate on real inputs
IF (fTotalTension <> fTotalTension) OR (fFrictionDrop <> fFrictionDrop)
   OR (fAccel <> fAccel) OR (fMassPerLen <> fMassPerLen)
   OR (ABS(fTotalTension) >= 3.0E38) OR (ABS(fFrictionDrop) >= 3.0E38)
   OR (ABS(fAccel) >= 3.0E38) OR (ABS(fMassPerLen) >= 3.0E38) THEN
    uErrorId := 16#0002_9226;   // 入参非有限拒收 / Non-finite input reject
    RETURN;
END_IF
// 段 2：域闸（根数下限防除零 + 摩擦/线密度非负，R4）/ Domain gate
IF iStrandCount < 1 THEN
    uErrorId := 16#0002_9226;   // 根数不足 1，单束张力不可解 / Strand count below one
    RETURN;
END_IF
IF (fFrictionDrop < 0.0) OR (fMassPerLen < 0.0) THEN
    uErrorId := 16#0002_9226;   // 摩擦损失或线密度为负 / Negative friction or density
    RETURN;
END_IF
// 段 3：主计算（有效总张力 → 单束张力 → cN）/ Main computation
fEffective := fTotalTension - fFrictionDrop + fMassPerLen * fAccel;     // 有效总张力 [N] / Effective tension
IF fEffective <= 1.0E-6 THEN
    uErrorId := 16#0002_9226;   // 有效总张力非正，物理不可达 / Effective tension non-positive
    RETURN;
END_IF
fTensionPerStrand := fEffective / INT_TO_REAL(iStrandCount) * 100.0;    // 单束张力 [cN] / Per strand
// 段 4：出口闸（非有限复核 + 正数复核）/ Outlet gate
IF (fTensionPerStrand <> fTensionPerStrand) OR (ABS(fTensionPerStrand) >= 3.0E38)
   OR (fTensionPerStrand <= 0.0) THEN
    fTensionPerStrand := 0.0;   // 复核失败回缺省 / Fallback on recheck failure
    uErrorId := 16#0002_9226;   // 出口复核拒收 / Output recheck reject
    RETURN;
END_IF
bValid := TRUE;                 // 有效回执 / Validity receipt
FC_DL_StrandTensionAtWinderCalc := fTensionPerStrand;   // 返回值镜像单束张力 / Return mirrors tension
END_FUNCTION

(* ---- FC_DL_StripCrownCalc.st ---- *)
(*
  Name: FC_DL_StripCrownCalc
  Category: DL_Device
  Version: 1.0.0
  Round: R89 / 2026-11-25
  开源溯源：clean-room 自研（族 板带剪切分条卷取，ST 开源生态实测 0 命中，无外部代码引入）
  功能：板凸度与平直度指数：由中部/边部厚度差算凸度（μm）、凸度率与 I-unit 平直度。
  边界条件：① 四入参全部过非有限闸，任一非有限返回哨兵 -1；
            ② 边部厚度为凸度率除子，须 ≥ 0.05 mm；凸度差取中部减边部，允许负值（负凸度照实输出）；
            ③ 平直度按「凸度差 ÷ 半宽」的应变 × 1e5 折算 I-unit，半宽为除子，带宽须 ≥ 200 mm；
            ④ fRefCrownPct 仅作域闸用的目标凸度率基准（0.1~5 %），不参与输出计算。
  量纲自证：(中部−边部)[mm]×1000 = μm；Δmm/(W/2)[mm] 无量纲 ×1e5 = I-unit。
*)
FUNCTION FC_DL_StripCrownCalc : REAL
VAR_INPUT
    fCenterThkMm : REAL;    (* 中部厚度 [mm] Center thickness [mm] *)
    fEdgeThkMm : REAL;      (* 边部厚度（距边 25 mm 处） [mm] Edge thickness [mm] *)
    fWidthMm : REAL;        (* 带钢宽度 [mm] Strip width [mm] *)
    fRefCrownPct : REAL;    (* 目标凸度率（域闸基准） [%] Reference crown ratio [%] *)
END_VAR
VAR_OUTPUT
    fCrownUm : REAL;        (* 凸度（中部−边部） [μm] Crown in micrometres [um] *)
    fCrownPct : REAL;       (* 凸度率（相对边部厚度） [%] Crown ratio [%] *)
    fFlatnessIu : REAL;     (* 平直度指数 [I-unit] Flatness index [I-unit] *)
    xValid : BOOL;          (* 计算有效性标志 [-] Calculation valid flag *)
END_VAR
VAR CONSTANT
    DL_EPS : REAL := 1.0E-9;        (* 判据容差 [-] Criterion tolerance *)
    DL_UM : REAL := 1000.0;         (* 毫米 → 微米换算 [μm/mm] Millimetre to micrometre *)
    DL_IU : REAL := 1.0E5;          (* 应变 → I-unit 换算 [-] Strain to I-unit *)
    DL_HALF : REAL := 2.0;          (* 半宽除数 [-] Half-width divisor *)
    DL_PCT : REAL := 100.0;         (* 百分数基准 [%] Percent base *)
    DL_C_MIN : REAL := 0.05;        (* 厚度下限 [mm] Thickness floor [mm] *)
    DL_C_MAX : REAL := 12.0;        (* 厚度上限 [mm] Thickness ceiling [mm] *)
    DL_W_MIN : REAL := 200.0;       (* 带宽下限 [mm] Width floor [mm] *)
    DL_W_MAX : REAL := 2500.0;      (* 带宽上限 [mm] Width ceiling [mm] *)
    DL_R_MIN : REAL := 0.1;         (* 目标凸度率下限 [%] Reference ratio floor [%] *)
    DL_R_MAX : REAL := 5.0;         (* 目标凸度率上限 [%] Reference ratio ceiling [%] *)
END_VAR
VAR
    fCrownMm : REAL;    (* 凸度差（mm） [mm] Crown difference [mm] *)
END_VAR
(* 出口预置：四出口统一预置（R256） *)
fCrownUm := 0.0; fCrownPct := 0.0; fFlatnessIu := 0.0; xValid := FALSE;
(* 非有限闸：NaN 自反判 + Inf 差值自减判，四入参全枚举 *)
IF (fCenterThkMm <> fCenterThkMm) OR ((fCenterThkMm - fCenterThkMm) <> 0.0)
   OR (fEdgeThkMm <> fEdgeThkMm) OR ((fEdgeThkMm - fEdgeThkMm) <> 0.0)
   OR (fWidthMm <> fWidthMm) OR ((fWidthMm - fWidthMm) <> 0.0)
   OR (fRefCrownPct <> fRefCrownPct) OR ((fRefCrownPct - fRefCrownPct) <> 0.0) THEN
    FC_DL_StripCrownCalc := -1.0;           (* 哨兵 -1：入参非有限 / Sentinel -1, non-finite input *)
    RETURN;
END_IF
(* 组态域闸：两侧厚度、带宽、目标凸度率逐项定域（边厚为凸度率除子） *)
IF (fCenterThkMm < DL_C_MIN) OR (fCenterThkMm > DL_C_MAX)
   OR (fEdgeThkMm < DL_C_MIN) OR (fEdgeThkMm > DL_C_MAX)
   OR (fWidthMm < DL_W_MIN) OR (fWidthMm > DL_W_MAX)
   OR (fRefCrownPct < DL_R_MIN) OR (fRefCrownPct > DL_R_MAX) THEN
    FC_DL_StripCrownCalc := -1.0;           (* 哨兵 -1：组态非法 / Sentinel -1, bad configuration *)
    RETURN;
END_IF
(* 凸度差：中部 − 边部，允许负值（负凸度照实上报，不做单向钳位） *)
fCrownMm := fCenterThkMm - fEdgeThkMm;
(* 凸度：mm × 1000 = μm *)
fCrownUm := fCrownMm * DL_UM;
(* 凸度率：÷ 边部厚度（已过下限闸），×100 得百分数 *)
fCrownPct := (fCrownMm / fEdgeThkMm) * DL_PCT;
(* 平直度：Δmm ÷ 半宽[mm] 得应变，×1e5 得 I-unit；半宽 = W/2 > 100 mm 恒正 *)
fFlatnessIu := (fCrownMm / (fWidthMm / DL_HALF)) * DL_IU;
xValid := TRUE;                             (* 链路有效 / Chain valid *)
FC_DL_StripCrownCalc := fCrownUm;
END_FUNCTION

(* ---- FC_DL_StripLengthAccumCalc.st ---- *)
(*
  Name: FC_DL_StripLengthAccumCalc
  Category: DL_Device
  Version: 1.0.0
  Round: R89 / 2026-11-25
  开源溯源：clean-room 自研（族 板带剪切分条卷取，ST 开源生态实测 0 命中，无外部代码引入）
  功能：带长累计：编码器脉冲差分解算 + 辊径磨损补偿，累积为米制长度。
  边界条件：① 两浮点入参过非有限闸，配置越域置 xValid = FALSE 并保持末值（不清零，防长度跳变）；
            ② 差分为负视为计数器清零或回绕：本拍不计入（reset 语义），并把快照更新到当前值；
            ③ 本件在 FC 内使用 VAR 保持量（上一拍脉冲、累计长度）；交付门槛：须在 CODESYS / TwinCAT /
               InoProShop 三平台各编译验证一次，确认 FC 局部静态量保留语义一致（R64 门槛声明）；
            ④ 有效辊径 = 标称辊径 − 磨损量，须 > 10 mm 否则判配置非法（周长为除数量纲基准）。
  量纲自证：脉冲数/每转脉冲数 = 转；转 × π·D[m] = m；D 由 mm/1000 得 m。
*)
FUNCTION FC_DL_StripLengthAccumCalc : REAL
VAR_INPUT
    nPulse : DINT;          (* 编码器累计脉冲（有符号，允许回绕） [pulse] Encoder pulse count [pulse] *)
    nPulsePerRev : DINT;    (* 每转脉冲数 [pulse/rev] Pulses per revolution [pulse/rev] *)
    fRollDiaMm : REAL;      (* 测量辊标称直径 [mm] Measuring roll nominal diameter [mm] *)
    fRollWearMm : REAL;     (* 测量辊累计磨损量 [mm] Roll accumulated wear [mm] *)
    xReset : BOOL;          (* 长度清零（换卷时置位一拍） [-] Reset accumulated length *)
END_VAR
VAR_OUTPUT
    fLengthM : REAL;        (* 累计长度 [m] Accumulated length [m] *)
    fRollDiaEffMm : REAL;   (* 有效（磨损后）辊径 [mm] Effective roll diameter [mm] *)
    xValid : BOOL;          (* 配置与链路有效 [-] Configuration and chain valid *)
END_VAR
VAR
    _nPulsePrev : DINT := 0;    (* 上一拍脉冲快照 [pulse] Previous pulse snapshot [pulse] *)
    _diDelta : DINT := 0;       (* 本拍脉冲增量 [pulse] Pulse increment [pulse] *)
    _fLenAccM : REAL := 0.0;    (* 累计长度保持量 [m] Accumulated length hold [m] *)
    _fCircM : REAL := 0.0;      (* 有效周长 [m] Effective circumference [m] *)
    _fDiaEff : REAL := 0.0;     (* 有效辊径保持量 [mm] Effective diameter hold [mm] *)
    _bCfgBad : BOOL := FALSE;   (* 配置非法当拍量 [-] Configuration bad *)
END_VAR
VAR CONSTANT
    DL_MM_TO_M : REAL := 1000.0;    (* 毫米 → 米换算 [mm/m] Millimetre to metre *)
    DL_DIA_MIN : REAL := 10.0;      (* 有效辊径下限 [mm] Effective diameter floor [mm] *)
    DL_DIA_MAX : REAL := 2000.0;    (* 标称辊径上限 [mm] Nominal diameter ceiling [mm] *)
    DL_WEAR_MAX : REAL := 50.0;     (* 磨损量上限 [mm] Wear ceiling [mm] *)
END_VAR
(* 出口预置：三出口与返回值统一预置（R256） *)
fLengthM := 0.0; fRollDiaEffMm := 0.0; xValid := FALSE; FC_DL_StripLengthAccumCalc := 0.0;
(* 非有限闸：NaN 自反判 + Inf 差值自减判，两浮点入参全枚举 *)
IF (fRollDiaMm <> fRollDiaMm) OR ((fRollDiaMm - fRollDiaMm) <> 0.0)
   OR (fRollWearMm <> fRollWearMm) OR ((fRollWearMm - fRollWearMm) <> 0.0) THEN
    fLengthM := _fLenAccM;                  (* 保持末值 / Hold last value *)
    fRollDiaEffMm := _fDiaEff;
    FC_DL_StripLengthAccumCalc := _fLenAccM;
    RETURN;
END_IF
(* 组态域闸：每转脉冲数为除子，磨损量不得吞掉辊径 *)
_bCfgBad := (nPulsePerRev < 1) OR (fRollDiaMm < (DL_DIA_MIN + DL_DIA_MIN))
         OR (fRollDiaMm > DL_DIA_MAX) OR (fRollWearMm < 0.0) OR (fRollWearMm > DL_WEAR_MAX);
IF _bCfgBad THEN
    fLengthM := _fLenAccM;                  (* 冻结保持，xValid 置假 / Freeze and mark invalid *)
    fRollDiaEffMm := _fDiaEff;
    FC_DL_StripLengthAccumCalc := _fLenAccM;
    RETURN;
END_IF
(* 有效辊径与周长：周长 = π·D，D 用米 *)
_fDiaEff := fRollDiaMm - fRollWearMm;
IF _fDiaEff <= DL_DIA_MIN THEN
    fLengthM := _fLenAccM;                  (* 磨损过限：冻结保持 / Wear too large, freeze *)
    fRollDiaEffMm := _fDiaEff;
    FC_DL_StripLengthAccumCalc := _fLenAccM;
    RETURN;
END_IF
_fCircM := 3.141592653589793 * (_fDiaEff / DL_MM_TO_M);
(* 脉冲差分：负增量视为计数器清零/回绕，本拍不计入 *)
_diDelta := nPulse - _nPulsePrev;
IF _diDelta > 0 THEN
    (* 转数 = 脉冲 ÷ 每转脉冲，再乘周长得米 *)
    _fLenAccM := _fLenAccM + (DINT_TO_REAL(_diDelta) / DINT_TO_REAL(nPulsePerRev)) * _fCircM;
END_IF
(* 清零：只清长度累计，不动配置（作用域声明） *)
IF xReset THEN
    _fLenAccM := 0.0;
END_IF
(* 末行更新快照：无论增量正负，快照都跟上，防回绕后重复计数 *)
_nPulsePrev := nPulse;
fLengthM := _fLenAccM;
fRollDiaEffMm := _fDiaEff;
xValid := TRUE;                             (* 链路有效 / Chain valid *)
FC_DL_StripLengthAccumCalc := fLengthM;
END_FUNCTION

(* ---- FC_DL_StripTensionRefCalc.st ---- *)
(*
  Name: FC_DL_StripTensionRefCalc
  Category: DL_Device
  Version: 1.0.0
  Round: R89 / 2026-11-25
  开源溯源：clean-room 自研（族 板带剪切分条卷取，ST 开源生态实测 0 命中，无外部代码引入）
  功能：带钢张力设定：按断面面积与单位张力算总张力，并按设备张力上限钳位输出。
  边界条件：① 四入参全部过非有限闸，任一非有限返回哨兵 -1；
            ② 断面尺寸与单位张力按工程域闸限定（宽 100~2500 mm、厚 0.1~6 mm、单位张力 10~200 MPa）；
            ③ 钳位属量值饱和：xClamped = TRUE 表示设定被设备上限截断，xValid 仍为 TRUE（事实未伪造）。
  量纲自证：W[mm]/1000 × T[mm]/1000 = m2；m2 × σ[MPa = MN/m2] = MN = 1000 kN；故 ÷1000 得 kN。
*)
FUNCTION FC_DL_StripTensionRefCalc : REAL
VAR_INPUT
    fWidthMm : REAL;         (* 带钢宽度 [mm] Strip width [mm] *)
    fThkMm : REAL;           (* 带钢厚度 [mm] Strip thickness [mm] *)
    fUnitTensionMpa : REAL;  (* 单位张力 [MPa] Unit tension [MPa] *)
    fTensionMaxKN : REAL;    (* 设备张力上限 [kN] Equipment tension ceiling [kN] *)
END_VAR
VAR_OUTPUT
    fTensionKN : REAL;       (* 张力设定值 [kN] Tension setpoint [kN] *)
    xClamped : BOOL;         (* 已按上限钳位 [-] Clamped by ceiling *)
    xValid : BOOL;           (* 计算有效性标志 [-] Calculation valid flag *)
END_VAR
VAR CONSTANT
    DL_EPS : REAL := 1.0E-9;        (* 判据容差 [-] Criterion tolerance *)
    DL_MM_TO_M : REAL := 1000.0;    (* 毫米 → 米换算 [mm/m] Millimetre to metre *)
    DL_MN_TO_KN : REAL := 1000.0;   (* 兆牛 → 千牛换算 [kN/MN] Meganewton to kilonewton *)
    DL_W_MIN : REAL := 100.0;       (* 带宽下限 [mm] Width floor [mm] *)
    DL_W_MAX : REAL := 2500.0;      (* 带宽上限 [mm] Width ceiling [mm] *)
    DL_T_MIN : REAL := 0.1;         (* 带厚下限 [mm] Thickness floor [mm] *)
    DL_T_MAX : REAL := 6.0;         (* 带厚上限 [mm] Thickness ceiling [mm] *)
    DL_U_MIN : REAL := 10.0;        (* 单位张力下限 [MPa] Unit tension floor [MPa] *)
    DL_U_MAX : REAL := 200.0;       (* 单位张力上限 [MPa] Unit tension ceiling [MPa] *)
    DL_F_MIN : REAL := 1.0;         (* 设备上限下限 [kN] Equipment ceiling floor [kN] *)
    DL_F_MAX : REAL := 500.0;       (* 设备上限上限 [kN] Equipment ceiling top [kN] *)
END_VAR
VAR
    fAreaM2 : REAL;     (* 断面面积 [m2] Cross-section area [m2] *)
    fForceMN : REAL;    (* 张力（兆牛） [MN] Tension in meganewtons [MN] *)
END_VAR
(* 出口预置：三出口统一预置（R256） *)
fTensionKN := 0.0; xClamped := FALSE; xValid := FALSE;
(* 非有限闸：NaN 自反判 + Inf 差值自减判，四入参全枚举 *)
IF (fWidthMm <> fWidthMm) OR ((fWidthMm - fWidthMm) <> 0.0)
   OR (fThkMm <> fThkMm) OR ((fThkMm - fThkMm) <> 0.0)
   OR (fUnitTensionMpa <> fUnitTensionMpa) OR ((fUnitTensionMpa - fUnitTensionMpa) <> 0.0)
   OR (fTensionMaxKN <> fTensionMaxKN) OR ((fTensionMaxKN - fTensionMaxKN) <> 0.0) THEN
    FC_DL_StripTensionRefCalc := -1.0;      (* 哨兵 -1：入参非有限 / Sentinel -1, non-finite input *)
    RETURN;
END_IF
(* 组态域闸：断面与单位张力、设备上限逐项定域 *)
IF (fWidthMm < DL_W_MIN) OR (fWidthMm > DL_W_MAX)
   OR (fThkMm < DL_T_MIN) OR (fThkMm > DL_T_MAX)
   OR (fUnitTensionMpa < DL_U_MIN) OR (fUnitTensionMpa > DL_U_MAX)
   OR (fTensionMaxKN < DL_F_MIN) OR (fTensionMaxKN > DL_F_MAX) THEN
    FC_DL_StripTensionRefCalc := -1.0;      (* 哨兵 -1：组态非法 / Sentinel -1, bad configuration *)
    RETURN;
END_IF
(* 断面面积：mm → m 后相乘，量纲 m2 *)
fAreaM2 := (fWidthMm / DL_MM_TO_M) * (fThkMm / DL_MM_TO_M);
(* 张力：m2 × MPa = MN（1 MPa = 1 MN/m2），再折 kN *)
fForceMN := fAreaM2 * fUnitTensionMpa;
fTensionKN := fForceMN * DL_MN_TO_KN;
(* 上限钳位：量值饱和并置钳位标志，有效性不受影响 *)
IF fTensionKN > fTensionMaxKN THEN
    fTensionKN := fTensionMaxKN;
    xClamped := TRUE;
END_IF
IF fTensionKN < DL_EPS THEN
    fTensionKN := 0.0;                      (* 微负残差归零 / Negative residual to zero *)
END_IF
xValid := TRUE;                             (* 链路有效 / Chain valid *)
FC_DL_StripTensionRefCalc := fTensionKN;
END_FUNCTION

(* ---- FC_DL_StsCraneRailClampChk.st ---- *)
(*
 * FC_DL_StsCraneRailClampChk | C1 | DL_Device
 * 功能：夹轨器/顶轨器状态与联锁判定（命令-反馈一致性与轨道在位）       单位：xClampOk/xIllegal 为布尔，nFaultCode 为 INT 码位
 * 工况边界：仅判定静态组合，不持定时器（超时由调用方 FB 计时）；xAnchorFb 作为轨道在位的冗余反证（顶轨器伸出必然压轨）；无轨命令夹轨最危险，码位优先级最高
 * 代数值回代：xClampCmd=TRUE、xClampFb=TRUE、xRailPresent=TRUE、xAnchorFb=FALSE → xClampOk=TRUE、xIllegal=FALSE、nFaultCode=0（与 spec 判定式一致）
 * 开源溯源：clean-room 自研，未复制任何第三方代码（无外部来源）
 *)
FUNCTION FC_DL_StsCraneRailClampChk : BOOL
VAR_INPUT
    xClampCmd   : BOOL;              // 夹轨命令 | rail clamp command
    xClampFb    : BOOL;              // 夹轨到位反馈 | rail clamp engaged feedback
    xRailPresent: BOOL;              // 轨道在位检测 | rail presence detection
    xAnchorFb   : BOOL;              // 顶轨器/锚定销到位反馈 | jack or anchor pin engaged feedback
END_VAR
VAR_OUTPUT
    xClampOk   : BOOL;               // 夹轨有效（命令+反馈+轨道三者成立）| clamp effective, command and feedback and rail
    xIllegal   : BOOL;               // 联锁非法 | interlock violation
    nFaultCode : INT;                // 0=无 / 9202=命令反馈不一致 / 9203=无轨夹轨 | 0 none, 9202 command-feedback mismatch, 9203 clamping without rail
    xRailOk    : BOOL;               // 轨道在位判定结果（含顶轨器冗余反证）| rail verdict including the jack redundancy
    xValid     : BOOL;               // 输出有效（无联锁非法）| outputs valid, no interlock violation
END_VAR

// 段1｜轨道在位：直接检测 OR 顶轨器到位反证（两个独立来源任一生效即认为在位）
xRailOk := xRailPresent OR xAnchorFb;

// 段2｜夹轨有效：命令、到位反馈、轨道三者同时成立
xClampOk := xClampCmd AND xClampFb AND xRailOk;

// 段3｜联锁非法判定（按危险度排序：无轨夹轨优先于命令反馈不一致）
xIllegal := FALSE;
nFaultCode := 0;
IF xClampCmd AND (NOT xRailOk) THEN
    xIllegal := TRUE;
    nFaultCode := 9203;              // 无轨夹轨：机构空夹，最危险 | clamping without a rail, the most dangerous case
ELSIF xClampCmd AND (NOT xClampFb) THEN
    xIllegal := TRUE;
    nFaultCode := 9202;              // 命令已给但未到位（由调用方 FB 计时判超时）| command given but not engaged, timed by the caller
ELSIF (NOT xClampCmd) AND xClampFb THEN
    xIllegal := TRUE;
    nFaultCode := 9202;              // 无命令却有到位反馈（反馈粘连或指令丢失）| feedback stuck on without a command
END_IF

// 段4｜出口
xValid := NOT xIllegal;
FC_DL_StsCraneRailClampChk := xValid;
END_FUNCTION

(* ---- FC_DL_SuctionCupCountCalc.st ---- *)
(*
  ============================================================
  组件名 : FC_DL_SuctionCupCountCalc
  分类   : DL_Device
  功能   : 吸盘数量配置计算，按载荷重力与冗余倾覆系数求所需吸盘数并给出可行性判定
  复杂度 : C2
  版本   : 1.0.0
  作者   : 道莅工业代码库工厂 / R81
  日期   : 2026-11-24
  开源溯源 : clean-room（no upstream）—— 依据公开工程公式自研，未复制任何上游实现
  红线自检 : R1 无GVL/R2 无物理地址/R3 纯IEC/R4 防除零/R5 双语注释
  接口说明 :
      需求数 = 向上取整(载荷kg * 9.81 * 冗余系数 * 倾覆系数 / 单盘可用力N)。
      向上取整不调用 CEIL，而是先截断再按余量进位，且截断前先做实数上限兜底，防止 REAL_TO_INT 溢出。
      结果限幅 1~64；需求数超过 32 时可行性判 FALSE，表示超出常规单机吸盘阵列规模。
      需求数溢出上限时直接按 64 落定并判不可行，不做回绕。
  ============================================================
*)
FUNCTION FC_DL_SuctionCupCountCalc : BOOL
VAR_INPUT
    bEnable      : BOOL; // 使能：TRUE 时计算 / Enable: TRUE to compute
    bErr         : BOOL; // 外部故障：TRUE 时立即退出并置结果无效 / External fault: TRUE aborts with invalid result
    rLoadKg      : REAL; // 被吸持工件质量 [kg] / mass of the workpiece to be held [kilogram]
    rPerCupN     : REAL; // 单个吸盘可用吸附力 [N] / usable holding force of one cup [newton]
    rRedundancy  : REAL; // 冗余系数，常用 1.2~2.0 [无量纲] / redundancy factor, typically 1.2 to 2.0 [dimensionless]
    rTiltFactor  : REAL; // 倾覆与动态系数 [无量纲] / tilt and dynamic factor [dimensionless]
END_VAR
VAR_OUTPUT
    rNeedRaw  : REAL; // 向上取整前的需求数 [个] / raw required count before rounding up [unit]
    iCupCnt   : INT;  // 配置吸盘数量，限幅 1~64 [个] / configured cup count clamped to 1 to 64 [unit]
    bFeasible : BOOL; // 可行：TRUE 表示数量不超过 32 个 / feasible, TRUE when the count does not exceed 32 [unit]
    bOverflow : BOOL; // 需求溢出：TRUE 表示需求数超出整数可表范围 / requirement overflow, TRUE when the requirement exceeds the integer range
    bValid    : BOOL; // 输出有效：TRUE 表示结果可用 / Output valid
END_VAR
VAR CONSTANT
    DL_R_MAX     : REAL := 3.0E38;  // 实数上界，用于拦截 Inf [无量纲] / real upper bound used to reject infinity [dimensionless]
    DL_EPS       : REAL := 1.0E-12; // 除零判定阈值 [无量纲] / division guard threshold [dimensionless]
    DL_G         : REAL := 9.81;    // 重力加速度 [m/s2] / gravitational acceleration [metre per second squared]
    DL_CUP_MIN   : INT := 1;        // 吸盘数量下界 [个] / lower bound of the cup count [unit]
    DL_CUP_MAX   : INT := 64;       // 吸盘数量上界 [个] / upper bound of the cup count [unit]
    DL_CUP_OK    : INT := 32;       // 常规阵列规模上限 [个] / upper bound of a conventional array [unit]
    DL_INT_SAFE  : REAL := 32000.0; // 实数转整数前的安全上限 [无量纲] / safe upper bound before converting a real into an integer [dimensionless]
    DL_RESID_TOL : REAL := 1.0E-6;  // 截断余量判定容差 [无量纲] / tolerance deciding the rounding carry [dimensionless]
    DL_RED_MIN   : REAL := 1.0;     // 冗余系数下界 [无量纲] / lower bound of the redundancy factor [dimensionless]
    DL_RED_MAX   : REAL := 5.0;     // 冗余系数上界 [无量纲] / upper bound of the redundancy factor [dimensionless]
    DL_TILT_MIN  : REAL := 1.0;     // 倾覆系数下界 [无量纲] / lower bound of the tilt factor [dimensionless]
    DL_TILT_MAX  : REAL := 5.0;     // 倾覆系数上界 [无量纲] / upper bound of the tilt factor [dimensionless]
    DL_LOAD_MAX  : REAL := 100000.0; // 工件质量合理上限 [kg] / sanity upper bound of the workpiece mass [kilogram]
END_VAR
VAR
    _bFin  : BOOL := FALSE; // 输入有限性判定结果 / input finiteness verdict
    _iTmp  : INT := 0;      // 截断后的临时整数 [个] / temporary integer after truncation [unit]
    _rRes  : REAL := 0.0;   // 截断余量 [个] / residual after truncation [unit]
END_VAR

    // 段 1｜出口预置：数量先置 1，可行位先置 FALSE
    rNeedRaw := 0.0;
    iCupCnt := DL_CUP_MIN;
    bFeasible := FALSE;
    bOverflow := FALSE;
    bValid := FALSE;
    // 段 2｜使能闸与外部故障闸
    IF NOT bEnable THEN
        RETURN;
    END_IF;
    IF bErr THEN
        RETURN;
    END_IF;
    // 段 3｜非有限闸
    _bFin := (rLoadKg = rLoadKg) AND (ABS(rLoadKg) <= DL_R_MAX) AND (rPerCupN = rPerCupN) AND (ABS(rPerCupN) <= DL_R_MAX) AND (rRedundancy = rRedundancy) AND (ABS(rRedundancy) <= DL_R_MAX) AND (rTiltFactor = rTiltFactor) AND (ABS(rTiltFactor) <= DL_R_MAX);
    IF NOT _bFin THEN
        RETURN;
    END_IF;
    // 段 4｜域闸：单盘力严格为正，载荷非负且合理，两个系数落在工程区间
    IF (ABS(rPerCupN) <= DL_EPS) OR (rPerCupN < 0.0) THEN
        RETURN;
    END_IF;
    IF (rLoadKg < 0.0) OR (rLoadKg > DL_LOAD_MAX) THEN
        RETURN;
    END_IF;
    IF (rRedundancy < DL_RED_MIN) OR (rRedundancy > DL_RED_MAX) THEN
        RETURN;
    END_IF;
    IF (rTiltFactor < DL_TILT_MIN) OR (rTiltFactor > DL_TILT_MAX) THEN
        RETURN;
    END_IF;
    // 段 5｜需求数原值
    rNeedRaw := rLoadKg * DL_G * rRedundancy * rTiltFactor / rPerCupN;
    // 段 6｜临界零需求：无载荷时按最小 1 个配置，直接判定
    IF rNeedRaw <= DL_RESID_TOL THEN
        iCupCnt := DL_CUP_MIN;
        bFeasible := TRUE;
        bOverflow := FALSE;
        bValid := TRUE;
        FC_DL_SuctionCupCountCalc := bValid;
        RETURN;
    END_IF;
    // 段 7｜实数上限兜底：超界直接按上界落定并判不可行，杜绝 REAL_TO_INT 回头
    IF rNeedRaw >= DL_INT_SAFE THEN
        iCupCnt := DL_CUP_MAX;
        bFeasible := FALSE;
        bOverflow := TRUE;
        bValid := TRUE;
        FC_DL_SuctionCupCountCalc := bValid;
        RETURN;
    END_IF;
    // 段 8｜先截断再按余量进位，等价向上取整但不调用 CEIL
    _iTmp := REAL_TO_INT(rNeedRaw);
    _rRes := rNeedRaw - INT_TO_REAL(_iTmp);
    IF _rRes > DL_RESID_TOL THEN
        _iTmp := _iTmp + 1;
    END_IF;
    // 段 9｜限幅与可行性
    IF _iTmp < DL_CUP_MIN THEN
        _iTmp := DL_CUP_MIN;
    END_IF;
    IF _iTmp > DL_CUP_MAX THEN
        _iTmp := DL_CUP_MAX;
    END_IF;
    iCupCnt := _iTmp;
    IF _iTmp <= DL_CUP_OK THEN
        bFeasible := TRUE;
    ELSE
        bFeasible := FALSE;
    END_IF;
    bOverflow := FALSE;
    bValid := TRUE;
    FC_DL_SuctionCupCountCalc := bValid;
END_FUNCTION

(* ---- FC_DL_SuctionFlowEst.st ---- *)
(*
  ============================================================
  组件名 : FC_DL_SuctionFlowEst
  分类   : DL_Device
  功能   : 真空抽吸流量估算，按喷嘴直径真空度与流量系数求可达到的抽吸体积流量
  复杂度 : C2
  版本   : 1.0.0
  作者   : 道莅工业代码库工厂 / R81
  日期   : 2026-11-24
  开源溯源 : clean-room（no upstream）—— 依据公开工程公式自研，未复制任何上游实现
  红线自检 : R1 无GVL/R2 无物理地址/R3 纯IEC/R4 防除零/R5 双语注释
  接口说明 :
      孔口流量式 Q = Cd * (pi/4) * (直径/1000)^2 * SQRT(2*压差/密度)，压差由 kPa 折 Pa，密度取 1.2 kg/m3。
      Q 的自然单位为 m3/s，乘以 60000/1000 即乘 60 后得到 L/min。
      该式为不可压缩孔口近似，仅在压比不进入临界区时可用，属工程估算而非精确标定。
  ============================================================
*)
FUNCTION FC_DL_SuctionFlowEst : BOOL
VAR_INPUT
    bEnable  : BOOL; // 使能：TRUE 时计算 / Enable: TRUE to compute
    bErr     : BOOL; // 外部故障：TRUE 时立即退出并置结果无效 / External fault: TRUE aborts with invalid result
    rDia_mm  : REAL; // 抽吸喷嘴等效直径 [mm] / equivalent nozzle diameter [millimetre]
    rVacKpa  : REAL; // 工作真空度 [kPa] / working vacuum level [kilopascal]
    rCd      : REAL; // 流量系数，常用 0.6~0.85 [无量纲] / discharge coefficient, typically 0.6 to 0.85 [dimensionless]
END_VAR
VAR_OUTPUT
    rVel_ms   : REAL; // 孔口等效流速 [m/s] / equivalent orifice velocity [metre per second]
    rFlowLpm  : REAL; // 折算抽吸流量 [L/min] / equivalent suction flow [litre per minute]
    rFlowNm3h : REAL; // 折算标准状态流量 [Nm3/h] / equivalent normal flow [normal cubic metre per hour]
    bValid    : BOOL; // 输出有效：TRUE 表示结果可用 / Output valid
END_VAR
VAR CONSTANT
    DL_PI       : REAL := 3.14159265; // 圆周率 [无量纲] / circular constant [dimensionless]
    DL_R_MAX    : REAL := 3.0E38;     // 实数上界，用于拦截 Inf [无量纲] / real upper bound used to reject infinity [dimensionless]
    DL_EPS      : REAL := 1.0E-12;    // 除零判定阈值 [无量纲] / division guard threshold [dimensionless]
    DL_MM_TO_M  : REAL := 1000.0;     // 毫米折米系数 [mm/m] / millimetre to metre factor [millimetre per metre]
    DL_KPA_TO_PA : REAL := 1000.0;    // 千帕折帕系数 [Pa/kPa] / kilopascal to pascal factor [pascal per kilopascal]
    DL_RHO      : REAL := 1.2;        // 空气密度 [kg/m3] / air density [kilogram per cubic metre]
    DL_QUARTER  : REAL := 0.25;       // 四分之一，用于 pi/4 折算 [无量纲] / one quarter used for the pi over four term [dimensionless]
    DL_M3S_TO_LPM : REAL := 60000.0;  // 立方米每秒折升每分系数（含 1/1000 体积换算）[无量纲] / cubic metre per second to litre per minute factor [dimensionless]
    DL_M3S_TO_NM3H : REAL := 3600.0;  // 立方米每秒折立方米每小时系数 [无量纲] / cubic metre per second to cubic metre per hour factor [dimensionless]
    DL_CD_MIN   : REAL := 0.1;        // 流量系数可信下界 [无量纲] / credible lower bound of the discharge coefficient [dimensionless]
    DL_CD_MAX   : REAL := 1.0;        // 流量系数物理上界 [无量纲] / physical upper bound of the discharge coefficient [dimensionless]
    DL_VAC_MAX  : REAL := 101.3;      // 真空度物理上限，标准大气压 [kPa] / physical upper bound of the vacuum level, standard atmosphere [kilopascal]
    DL_DIA_MAX  : REAL := 1000.0;     // 喷嘴直径合理上限 [mm] / sanity upper bound of the nozzle diameter [millimetre]
END_VAR
VAR
    _bFin  : BOOL := FALSE; // 输入有限性判定结果 / input finiteness verdict
    _rDia  : REAL := 0.0;   // 喷嘴直径折算米 [m] / nozzle diameter in metre [metre]
    _rArea : REAL := 0.0;   // 喷嘴过流面积 [m2] / nozzle flow area [square metre]
    _rPress : REAL := 0.0;  // 压差折算帕 [Pa] / differential pressure in pascal [pascal]
    _rTerm : REAL := 0.0;   // 流速根号内被开方数 [m2/s2] / radicand of the velocity square root [square metre per square second]
    _rQm3s : REAL := 0.0;   // 体积流量 [m3/s] / volumetric flow [cubic metre per second]
END_VAR

    // 段 1｜出口预置
    rVel_ms := 0.0;
    rFlowLpm := 0.0;
    rFlowNm3h := 0.0;
    bValid := FALSE;
    // 段 2｜使能闸与外部故障闸
    IF NOT bEnable THEN
        RETURN;
    END_IF;
    IF bErr THEN
        RETURN;
    END_IF;
    // 段 3｜非有限闸
    _bFin := (rDia_mm = rDia_mm) AND (ABS(rDia_mm) <= DL_R_MAX) AND (rVacKpa = rVacKpa) AND (ABS(rVacKpa) <= DL_R_MAX) AND (rCd = rCd) AND (ABS(rCd) <= DL_R_MAX);
    IF NOT _bFin THEN
        RETURN;
    END_IF;
    // 段 4｜域闸
    IF (ABS(rDia_mm) <= DL_EPS) OR (rDia_mm < 0.0) OR (rDia_mm > DL_DIA_MAX) THEN
        RETURN;
    END_IF;
    IF (ABS(rVacKpa) <= DL_EPS) OR (rVacKpa < 0.0) OR (rVacKpa > DL_VAC_MAX) THEN
        RETURN;
    END_IF;
    IF (rCd < DL_CD_MIN) OR (rCd > DL_CD_MAX) THEN
        RETURN;
    END_IF;
    // 段 5｜面积与压差
    _rDia := rDia_mm / DL_MM_TO_M;
    _rArea := DL_PI * DL_QUARTER * _rDia * _rDia;
    _rPress := rVacKpa * DL_KPA_TO_PA;
    // 段 6｜开方前必须确认被开方数非负，密度分母已按常数保证为正
    _rTerm := 2.0 * _rPress / DL_RHO;
    IF _rTerm < 0.0 THEN
        RETURN;
    END_IF;
    rVel_ms := SQRT(_rTerm);
    // 段 7｜体积流量与单位折算
    _rQm3s := rCd * _rArea * rVel_ms;
    rFlowLpm := _rQm3s * DL_M3S_TO_LPM;
    rFlowNm3h := _rQm3s * DL_M3S_TO_NM3H;
    bValid := TRUE;
    FC_DL_SuctionFlowEst := bValid;
END_FUNCTION

(* ---- FC_DL_ToolWearVbCalc.st ---- *)
(*
  DL Factory R84 | FC_DL_ToolWearVbCalc
  功能：按磨损速率算后刀面磨损量 VB 与到磨损限值的剩余可用时间
  开源溯源：无（clean-room 自研，依据公开工艺公式，来源=行业通用公式，许可证=MIT，借鉴点=公式结构）
  规则：R1-R16 全遵守
*)
FUNCTION FC_DL_ToolWearVbCalc : REAL
VAR_INPUT
    fVb0Mm : REAL := 0.05; // 初始后刀面磨损 [mm] / initial flank wear [mm]
    fKMmPerM : REAL := 0.00002; // 磨损系数（每米切削路程增量） [mm/m] / wear coefficient [mm/m]
    fVcMpm : REAL := 200.0; // 切削线速度 [m/min] / cutting speed [m/min]
    fTimeMin : REAL := 10.0; // 累计切削时间 [min] / accumulated cutting time [min]
    fVbLimitMm : REAL := 0.30; // 后刀面磨损限值（换刀判据） [mm] / flank wear limit [mm]
END_VAR
VAR_OUTPUT
    fRemainMin : REAL; // 到限值剩余可用时间 [min] / remaining usable time [min]
    xWorn : BOOL; // 已达磨损限值 [-] / wear limit reached [-]
    xValid : BOOL; // 计算结果有效标志 [-] / calculation valid flag [-]
END_VAR
VAR
    fPathM : REAL; // 累计切削路程 [m] / accumulated cutting path [m]
    fVbRaw : REAL; // 磨损量中间量 [mm] / wear intermediate [mm]
    fRateMmPerMin : REAL; // 磨损速率 [mm/min] / wear rate [mm/min]
END_VAR

// 段 1｜出口预置（R256）
FC_DL_ToolWearVbCalc := -1.0; // 哨兵返回 -1（无效） [-] / sentinel return -1, invalid [-]
fRemainMin := 0.0; // 剩余时间预置零 [min] / remaining time preset zero [min]
xWorn := FALSE; // 磨损到位位预置 FALSE [-] / wear flag preset false [-]
xValid := FALSE; // 计算完成前不认结果 [-] / unusable before calculation [-]

// 段 2｜非有限拦截 + 域闸（R4/R20）
IF NOT (fVb0Mm > -1.0E30 AND fVb0Mm < 1.0E30) OR NOT (fKMmPerM > -1.0E30 AND fKMmPerM < 1.0E30) OR NOT (fVcMpm > -1.0E30 AND fVcMpm < 1.0E30) OR NOT (fTimeMin > -1.0E30 AND fTimeMin < 1.0E30) OR NOT (fVbLimitMm > -1.0E30 AND fVbLimitMm < 1.0E30) THEN
    RETURN; // 任一入参为 NaN/Inf 一律拒绝 [-] / any NaN or Inf input rejected [-]
END_IF
IF fVb0Mm < 0.0 OR fKMmPerM < 0.0 OR fVcMpm < 0.0 OR fTimeMin < 0.0 OR fVbLimitMm < 1.0E-9 THEN
    RETURN; // 磨损量/系数/速度/时间负域或限值非正即非法 [mm] / negative domains or non positive limit [mm]
END_IF

// 段 3｜VB = VB0 + k × (vc × t)
fPathM := fVcMpm * fTimeMin; // m/min × min = m / [m/min] × [min] = [m]
fVbRaw := fVb0Mm + (fKMmPerM * fPathM); // mm + mm/m × m = mm / [mm] + [mm/m] × [m] = [mm]
IF NOT (fVbRaw > -1.0E30 AND fVbRaw < 1.0E30) THEN
    RETURN; // 结果非有限再拦一次 [-] / second finiteness gate on the result [-]
END_IF

// 段 4｜剩余时间 = (限值 − VB) / 磨损速率
fRateMmPerMin := fKMmPerM * fVcMpm; // mm/m × m/min = mm/min / [mm/m] × [m/min] = [mm/min]
IF fVbRaw >= fVbLimitMm THEN
    xWorn := TRUE; // 已达/超限：剩余时间为零 [-] / limit reached, no remaining time [-]
    fRemainMin := 0.0; // 剩余时间钳零 [min] / clamp remaining time to zero [min]
ELSIF fRateMmPerMin < 1.0E-9 THEN
    fRemainMin := -1.0; // 分母闸：磨损速率趋零则剩余时间不可估 [min] / denominator gate, wear rate near zero [min]
ELSE
    fRemainMin := (fVbLimitMm - fVbRaw) / fRateMmPerMin; // mm ÷ mm/min = min / [mm] / [mm/min] = [min]
END_IF
xValid := TRUE; // 链路有效 [-] / chain valid [-]
FC_DL_ToolWearVbCalc := fVbRaw; // 返回磨损量 [mm] / return the flank wear [mm]
END_FUNCTION

(* ---- FC_DL_TurbidityNtuCalc.st ---- *)
(* ============================================================
   DL_Device / FC_DL_TurbidityNtuCalc ｜ v1.0.0 ｜ 2026-11-25
   功能：浊度比值法 ratio = (S − D) / (T − D)，NTU = K · ratio + Zero，
         末尾做负值保护与量程上限栅。
   边界：净透射 ≤ 1E-6（遮光/断线）或量程上限 ≤ 0 → 码 1、NTU 写 0（N1）；
         任一入参非有限 → 码 2、NTU 写 0；换算值为负 → 钳 0 报码 3；
         超量程上限 → 钳顶报码 4（饱和上报，值仍可读）。
         量纲清单（N5）：S/T/D 同一光路电压 [mV]，ratio 无量纲；K 单位 NTU/ratio；
         Zero 与上限同为 NTU；1 NTU = 1 FNU。
   依赖：仅 IEC 61131-3（无外部依赖，纯算术） ｜ 溯源：DLF-D-WATERANA
   验收：S=800/T=400/D=0/K=2.0/Zero=0.2/Max=1000 → ratio=2.0、NTU=4.2、码 0；
         T=0 → 码 1、NTU=0；结果超上限 → 钳顶、码 4。
   ============================================================ *)
FUNCTION FC_DL_TurbidityNtuCalc : BOOL
VAR_INPUT
    fScatterV  : REAL;  // 散射光路电压 [mV] / Scattered light channel voltage
    fTransmitV : REAL;  // 透射光路电压 [mV] / Transmitted light channel voltage
    fDarkV     : REAL;  // 暗电流（遮光）基准电压 [mV] / Dark current baseline voltage
    fKScale    : REAL;  // 标定系数，有效域 > 0 [NTU/ratio] / Calibration factor in NTU per ratio unit
    fZeroNtu   : REAL;  // 零点浊度偏置 [NTU] / Zero point turbidity offset
    fNtuMax    : REAL;  // 量程上限，有效域 > 0 [NTU] / Upper range limit of the measurement
END_VAR
VAR_OUTPUT
    fNtu   : REAL;   // 浊度换算值 [NTU] / Turbidity in nephelometric turbidity units
    uErrId : UDINT;  // 码 0 正常 / 1 遮光或组态非法 / 2 非有限 / 3 负值钳零 / 4 超量程钳顶 [-] / Outlet code
END_VAR
VAR
    _fS     : REAL;  // 净散射电压 [mV] / Net scattered light voltage
    _fT     : REAL;  // 净透射电压 [mV] / Net transmitted light voltage
    _fNtu   : REAL;  // 换算中间值 [NTU] / Intermediate turbidity value
END_VAR
VAR CONSTANT
    DL_TBN_EPS : REAL := 1.0E-6;  // 净透射判零下限 [mV] / Zero floor of the net transmitted voltage
END_VAR

(* 段 0：出口预置安全侧（0 NTU、码取最严，N1/N3） *)
FC_DL_TurbidityNtuCalc := FALSE;
fNtu := 0.0;  uErrId := 2;

(* 段 1：非有限闸（六个入参全量枚举；NaN 自反 + Inf 差值自减双判，R79/R272） *)
IF (fScatterV <> fScatterV) OR (fTransmitV <> fTransmitV) OR (fDarkV <> fDarkV)
   OR (fKScale <> fKScale) OR (fZeroNtu <> fZeroNtu) OR (fNtuMax <> fNtuMax) THEN RETURN; END_IF
(* Inf 双判须覆盖 fScatterV / fTransmitV / fDarkV：透射 +Inf 时净透射为 ±Inf，
   判零闸放行、比值算成 0，输出「NTU = Zero、码 0」的伪读数 *)
IF ((fScatterV - fScatterV) <> (fScatterV - fScatterV))
   OR ((fTransmitV - fTransmitV) <> (fTransmitV - fTransmitV))
   OR ((fDarkV - fDarkV) <> (fDarkV - fDarkV))
   OR ((fKScale - fKScale) <> (fKScale - fKScale))
   OR ((fZeroNtu - fZeroNtu) <> (fZeroNtu - fZeroNtu))
   OR ((fNtuMax - fNtuMax) <> (fNtuMax - fNtuMax)) THEN RETURN; END_IF

(* 段 2：域闸（净透射判零 + 系数与量程上限必须为正） *)
_fS := fScatterV - fDarkV;
_fT := fTransmitV - fDarkV;
IF (ABS(_fT) <= DL_TBN_EPS) OR (fKScale <= 0.0) OR (fNtuMax <= 0.0) THEN
    uErrId := 1;                        // 遮光/断线或组态非法：浊度不可解
    RETURN;
END_IF

(* 段 3：比值换算（除子已证 |T_net| > 1E-6） *)
_fNtu := fKScale * (_fS / _fT) + fZeroNtu;

(* 段 4：结果复检（非有限保持段 0 安全侧） *)
IF (_fNtu <> _fNtu) OR ((_fNtu - _fNtu) <> (_fNtu - _fNtu)) THEN RETURN; END_IF

(* 段 5：单一出口裁决（先钳后赋，判据与出口同源于 _fNtu，N4/R23） *)
IF _fNtu < 0.0 THEN
    fNtu := 0.0;  uErrId := 3;          // 负值保护：钳零后上报
ELSIF _fNtu > fNtuMax THEN
    fNtu := fNtuMax;  uErrId := 4;      // 饱和上报：钳顶后值仍可读
ELSE
    fNtu := _fNtu;  uErrId := 0;  FC_DL_TurbidityNtuCalc := TRUE;
END_IF
END_FUNCTION
